  MoveL 3592 to (0, -43.6, 16.44) mm, rotated rx 90 ry 0 rz 180 deg; joints [1.406, -71.721, 106.574, -177.541, 34.877, 177.982]
  MoveL 3593 to (0, -43.6, 17.04) mm, rotated rx 90 ry 0 rz 180 deg; joints [1.381, -71.722, 106.575, -177.584, 34.877, 178.018]
  MoveL 3594 to (-200, -43.6, 17.04) mm, rotated rx 90 ry 0 rz 180 deg; joints [1.617, -84.213, 122.025, -177.364, 37.842, 177.918]
  MoveL 3595 to (-200, -43.6, 17.64) mm, rotated rx 90 ry 0 rz 180 deg; joints [1.587, -84.214, 122.026, -177.412, 37.841, 177.956]
  MoveL 3596 to (0, -43.6, 17.64) mm, rotated rx 90 ry 0 rz 180 deg; joints [1.356, -71.723, 106.576, -177.628, 34.876, 178.054]
  MoveL 3597 to (0, -43.6, 18.24) mm, rotated rx 90 ry 0 rz 180 deg; joints [1.331, -71.724, 106.577, -177.672, 34.876, 178.09]
  MoveL 3598 to (-200, -43.6, 18.24) mm, rotated rx 90 ry 0 rz 180 deg; joints [1.558, -84.215, 122.027, -177.46, 37.84, 177.993]
  MoveL 3599 to (-200, -43.6, 18.84) mm, rotated rx 90 ry 0 rz 180 deg; joints [1.529, -84.216, 122.028, -177.508, 37.839, 178.031]
  MoveL 3600 to (0, -43.6, 18.84) mm, rotated rx 90 ry 0 rz 180 deg; joints [1.306, -71.725, 106.578, -177.716, 34.875, 178.126]
  MoveL 3601 to (0, -43.6, 19.44) mm, rotated rx 90 ry 0 rz 180 deg; joints [1.281, -71.725, 106.579, -177.759, 34.875, 178.162]
  MoveL 3602 to (-200, -43.6, 19.44) mm, rotated rx 90 ry 0 rz 180 deg; joints [1.499, -84.217, 122.03, -177.555, 37.838, 178.069]
  MoveL 3603 to (-200, -43.6, 20.04) mm, rotated rx 90 ry 0 rz 180 deg; joints [1.47, -84.218, 122.031, -177.603, 37.837, 178.107]
  MoveL 3604 to (0, -43.6, 20.04) mm, rotated rx 90 ry 0 rz 180 deg; joints [1.256, -71.726, 106.58, -177.803, 34.874, 178.197]
  MoveL 3605 to (0, -43.6, 20.64) mm, rotated rx 90 ry 0 rz 180 deg; joints [1.231, -71.727, 106.582, -177.847, 34.874, 178.233]
  MoveL 3606 to (-200, -43.6, 20.64) mm, rotated rx 90 ry 0 rz 180 deg; joints [1.441, -84.219, 122.032, -177.651, 37.836, 178.144]
  MoveL 3607 to (-200, -43.6, 21.24) mm, rotated rx 90 ry 0 rz 180 deg; joints [1.411, -84.22, 122.033, -177.699, 37.835, 178.182]
  MoveL 3608 to (0, -43.6, 21.24) mm, rotated rx 90 ry 0 rz 180 deg; joints [1.206, -71.728, 106.583, -177.891, 34.873, 178.269]
  MoveL 3609 to (0, -43.6, 21.84) mm, rotated rx 90 ry 0 rz 180 deg; joints [1.181, -71.729, 106.584, -177.935, 34.873, 178.305]
  MoveL 3610 to (-200, -43.6, 21.84) mm, rotated rx 90 ry 0 rz 180 deg; joints [1.382, -84.221, 122.034, -177.746, 37.835, 178.22]
  MoveL 3611 to (-200, -43.6, 22.44) mm, rotated rx 90 ry 0 rz 180 deg; joints [1.353, -84.222, 122.035, -177.794, 37.834, 178.258]
  MoveL 3612 to (0, -43.6, 22.44) mm, rotated rx 90 ry 0 rz 180 deg; joints [1.156, -71.729, 106.585, -177.978, 34.872, 178.341]
  MoveL 3613 to (0, -43.6, 23.04) mm, rotated rx 90 ry 0 rz 180 deg; joints [1.131, -71.73, 106.586, -178.022, 34.872, 178.377]
  MoveL 3614 to (-200, -43.6, 23.04) mm, rotated rx 90 ry 0 rz 180 deg; joints [1.323, -84.223, 122.036, -177.842, 37.833, 178.295]
  MoveL 3615 to (-200, -43.6, 23.64) mm, rotated rx 90 ry 0 rz 180 deg; joints [1.294, -84.223, 122.037, -177.89, 37.832, 178.333]
  MoveL 3616 to (0, -43.6, 23.64) mm, rotated rx 90 ry 0 rz 180 deg; joints [1.106, -71.731, 106.587, -178.066, 34.871, 178.413]
  MoveL 3617 to (0, -43.6, 24.24) mm, rotated rx 90 ry 0 rz 180 deg; joints [1.081, -71.731, 106.588, -178.11, 34.871, 178.449]
  MoveL 3618 to (-200, -43.6, 24.24) mm, rotated rx 90 ry 0 rz 180 deg; joints [1.265, -84.224, 122.038, -177.938, 37.832, 178.371]
  MoveL 3619 to (-200, -43.6, 24.84) mm, rotated rx 90 ry 0 rz 180 deg; joints [1.236, -84.225, 122.039, -177.985, 37.831, 178.408]
  MoveL 3620 to (0, -43.6, 24.84) mm, rotated rx 90 ry 0 rz 180 deg; joints [1.055, -71.732, 106.589, -178.154, 34.87, 178.485]
  MoveL 3621 to (0, -43.6, 25.44) mm, rotated rx 90 ry 0 rz 180 deg; joints [1.03, -71.733, 106.589, -178.197, 34.87, 178.521]
  MoveL 3622 to (-200, -43.6, 25.44) mm, rotated rx 90 ry 0 rz 180 deg; joints [1.206, -84.226, 122.04, -178.033, 37.83, 178.446]
  MoveL 3623 to (-200, -43.6, 26.04) mm, rotated rx 90 ry 0 rz 180 deg; joints [1.177, -84.227, 122.041, -178.081, 37.829, 178.484]
  MoveL 3624 to (0, -43.6, 26.04) mm, rotated rx 90 ry 0 rz 180 deg; joints [1.005, -71.733, 106.59, -178.241, 34.87, 178.557]
  MoveL 3625 to (0, -43.6, 26.64) mm, rotated rx 90 ry 0 rz 180 deg; joints [0.98, -71.734, 106.591, -178.285, 34.869, 178.593]
  MoveL 3626 to (-200, -43.6, 26.64) mm, rotated rx 90 ry 0 rz 180 deg; joints [1.148, -84.228, 122.042, -178.129, 37.829, 178.522]
  MoveL 3627 to (-200, -43.6, 27.24) mm, rotated rx 90 ry 0 rz 180 deg; joints [1.118, -84.228, 122.042, -178.176, 37.828, 178.559]
  MoveL 3628 to (0, -43.6, 27.24) mm, rotated rx 90 ry 0 rz 180 deg; joints [0.955, -71.735, 106.592, -178.329, 34.869, 178.629]
  MoveL 3629 to (0, -43.6, 27.84) mm, rotated rx 90 ry 0 rz 180 deg; joints [0.93, -71.735, 106.593, -178.373, 34.868, 178.665]
  MoveL 3630 to (-200, -43.6, 27.84) mm, rotated rx 90 ry 0 rz 180 deg; joints [1.089, -84.229, 122.043, -178.224, 37.827, 178.597]
  MoveL 3631 to (-200, -43.6, 28.44) mm, rotated rx 90 ry 0 rz 180 deg; joints [1.06, -84.23, 122.044, -178.272, 37.827, 178.635]
  MoveL 3632 to (0, -43.6, 28.44) mm, rotated rx 90 ry 0 rz 180 deg; joints [0.905, -71.736, 106.594, -178.417, 34.868, 178.701]
  MoveL 3633 to (0, -43.6, 29.04) mm, rotated rx 90 ry 0 rz 180 deg; joints [0.88, -71.737, 106.594, -178.46, 34.868, 178.737]
  MoveL 3634 to (-200, -43.6, 29.04) mm, rotated rx 90 ry 0 rz 180 deg; joints [1.03, -84.23, 122.045, -178.32, 37.826, 178.673]
  MoveL 3635 to (-200, -43.6, 29.64) mm, rotated rx 90 ry 0 rz 180 deg; joints [1.001, -84.231, 122.046, -178.368, 37.826, 178.711]
  MoveL 3636 to (0, -43.6, 29.64) mm, rotated rx 90 ry 0 rz 180 deg; joints [0.855, -71.737, 106.595, -178.504, 34.867, 178.773]
  MoveL 3637 to (0, -43.6, 30.24) mm, rotated rx 90 ry 0 rz 180 deg; joints [0.83, -71.738, 106.596, -178.548, 34.867, 178.809]
  MoveL 3638 to (-200, -43.6, 30.24) mm, rotated rx 90 ry 0 rz 180 deg; joints [0.972, -84.232, 122.046, -178.416, 37.825, 178.748]
  MoveL 3639 to (-200, -43.6, 30.84) mm, rotated rx 90 ry 0 rz 180 deg; joints [0.942, -84.232, 122.047, -178.463, 37.825, 178.786]
  MoveL 3640 to (0, -43.6, 30.84) mm, rotated rx 90 ry 0 rz 180 deg; joints [0.805, -71.738, 106.597, -178.592, 34.867, 178.845]
  MoveL 3641 to (0, -43.6, 31.44) mm, rotated rx 90 ry 0 rz 180 deg; joints [0.78, -71.739, 106.597, -178.636, 34.866, 178.88]
  MoveL 3642 to (-200, -43.6, 31.44) mm, rotated rx 90 ry 0 rz 180 deg; joints [0.913, -84.233, 122.048, -178.511, 37.824, 178.824]
  MoveL 3643 to (-200, -43.6, 32.04) mm, rotated rx 90 ry 0 rz 180 deg; joints [0.884, -84.234, 122.048, -178.559, 37.823, 178.862]
  MoveL 3644 to (0, -43.6, 32.04) mm, rotated rx 90 ry 0 rz 180 deg; joints [0.755, -71.739, 106.598, -178.679, 34.866, 178.916]
  MoveL 3645 to (0, -43.6, 32.64) mm, rotated rx 90 ry 0 rz 180 deg; joints [0.73, -71.74, 106.599, -178.723, 34.866, 178.952]
  MoveL 3646 to (-200, -43.6, 32.64) mm, rotated rx 90 ry 0 rz 180 deg; joints [0.854, -84.234, 122.049, -178.607, 37.823, 178.899]
  MoveL 3647 to (-200, -43.6, 33.24) mm, rotated rx 90 ry 0 rz 180 deg; joints [0.825, -84.235, 122.05, -178.655, 37.822, 178.937]
  MoveL 3648 to (0, -43.6, 33.24) mm, rotated rx 90 ry 0 rz 180 deg; joints [0.705, -71.74, 106.599, -178.767, 34.865, 178.988]
  MoveL 3649 to (0, -43.6, 33.84) mm, rotated rx 90 ry 0 rz 180 deg; joints [0.68, -71.741, 106.6, -178.811, 34.865, 179.024]
  MoveL 3650 to (-200, -43.6, 33.84) mm, rotated rx 90 ry 0 rz 180 deg; joints [0.796, -84.235, 122.05, -178.702, 37.822, 178.975]
  MoveL 3651 to (-200, -43.6, 34.44) mm, rotated rx 90 ry 0 rz 180 deg; joints [0.766, -84.236, 122.051, -178.75, 37.822, 179.013]
  MoveL 3652 to (0, -43.6, 34.44) mm, rotated rx 90 ry 0 rz 180 deg; joints [0.655, -71.741, 106.6, -178.855, 34.865, 179.06]
  MoveL 3653 to (0, -43.6, 35.04) mm, rotated rx 90 ry 0 rz 180 deg; joints [0.63, -71.741, 106.601, -178.899, 34.865, 179.096]
  MoveL 3654 to (-200, -43.6, 35.04) mm, rotated rx 90 ry 0 rz 180 deg; joints [0.737, -84.236, 122.051, -178.798, 37.821, 179.05]
  MoveL 3655 to (-200, -43.6, 35.64) mm, rotated rx 90 ry 0 rz 180 deg; joints [0.708, -84.237, 122.052, -178.846, 37.821, 179.088]
  MoveL 3656 to (0, -43.6, 35.64) mm, rotated rx 90 ry 0 rz 180 deg; joints [0.605, -71.742, 106.602, -178.942, 34.864, 179.132]
  MoveL 3657 to (0, -43.6, 36.24) mm, rotated rx 90 ry 0 rz 180 deg; joints [0.579, -71.742, 106.602, -178.986, 34.864, 179.168]
  MoveL 3658 to (-200, -43.6, 36.24) mm, rotated rx 90 ry 0 rz 180 deg; joints [0.678, -84.237, 122.053, -178.894, 37.82, 179.126]
  MoveL 3659 to (-200, -43.6, 36.84) mm, rotated rx 90 ry 0 rz 180 deg; joints [0.649, -84.238, 122.053, -178.942, 37.82, 179.164]
  MoveL 3660 to (0, -43.6, 36.84) mm, rotated rx 90 ry 0 rz 180 deg; joints [0.554, -71.743, 106.603, -179.03, 34.864, 179.204]
  MoveL 3661 to (0, -43.6, 37.44) mm, rotated rx 90 ry 0 rz 180 deg; joints [0.529, -71.743, 106.603, -179.074, 34.864, 179.24]
  MoveL 3662 to (-200, -43.6, 37.44) mm, rotated rx 90 ry 0 rz 180 deg; joints [0.62, -84.238, 122.053, -178.989, 37.82, 179.202]
  MoveL 3663 to (-200, -43.6, 38.04) mm, rotated rx 90 ry 0 rz 180 deg; joints [0.59, -84.239, 122.054, -179.037, 37.819, 179.239]
  MoveL 3664 to (0, -43.6, 38.04) mm, rotated rx 90 ry 0 rz 180 deg; joints [0.504, -71.743, 106.603, -179.118, 34.863, 179.276]
  MoveL 3665 to (0, -43.6, 38.64) mm, rotated rx 90 ry 0 rz 180 deg; joints [0.479, -71.744, 106.604, -179.162, 34.863, 179.312]
  MoveL 3666 to (-200, -43.6, 38.64) mm, rotated rx 90 ry 0 rz 180 deg; joints [0.561, -84.239, 122.054, -179.085, 37.819, 179.277]
  MoveL 3667 to (-200, -43.6, 39.24) mm, rotated rx 90 ry 0 rz 180 deg; joints [0.532, -84.239, 122.055, -179.133, 37.819, 179.315]
  MoveL 3668 to (0, -43.6, 39.24) mm, rotated rx 90 ry 0 rz 180 deg; joints [0.454, -71.744, 106.604, -179.205, 34.863, 179.348]
  MoveL 3669 to (0, -43.6, 39.84) mm, rotated rx 90 ry 0 rz 180 deg; joints [0.429, -71.744, 106.605, -179.249, 34.863, 179.384]
  MoveL 3670 to (-200, -43.6, 39.84) mm, rotated rx 90 ry 0 rz 180 deg; joints [0.502, -84.24, 122.055, -179.181, 37.818, 179.353]
  MoveL 3671 to (-200, -43.6, 40.44) mm, rotated rx 90 ry 0 rz 180 deg; joints [0.473, -84.24, 122.056, -179.229, 37.818, 179.391]
  MoveL 3672 to (0, -43.6, 40.44) mm, rotated rx 90 ry 0 rz 180 deg; joints [0.404, -71.744, 106.605, -179.293, 34.863, 179.42]
  MoveL 3673 to (0, -43.6, 41.04) mm, rotated rx 90 ry 0 rz 180 deg; joints [0.379, -71.745, 106.605, -179.337, 34.863, 179.456]
  MoveL 3674 to (-200, -43.6, 41.04) mm, rotated rx 90 ry 0 rz 180 deg; joints [0.444, -84.24, 122.056, -179.276, 37.818, 179.428]
  MoveL 3675 to (-200, -43.6, 41.64) mm, rotated rx 90 ry 0 rz 180 deg; joints [0.414, -84.241, 122.056, -179.324, 37.817, 179.466]
  MoveL 3676 to (0, -43.6, 41.64) mm, rotated rx 90 ry 0 rz 180 deg; joints [0.354, -71.745, 106.606, -179.381, 34.862, 179.492]
  MoveL 3677 to (0, -43.6, 42.24) mm, rotated rx 90 ry 0 rz 180 deg; joints [0.329, -71.745, 106.606, -179.425, 34.862, 179.528]
  MoveL 3678 to (-200, -43.6, 42.24) mm, rotated rx 90 ry 0 rz 180 deg; joints [0.385, -84.241, 122.057, -179.372, 37.817, 179.504]
  MoveL 3679 to (-200, -43.6, 42.84) mm, rotated rx 90 ry 0 rz 180 deg; joints [0.356, -84.241, 122.057, -179.42, 37.817, 179.542]
  MoveL 3680 to (0, -43.6, 42.84) mm, rotated rx 90 ry 0 rz 180 deg; joints [0.304, -71.745, 106.606, -179.468, 34.862, 179.564]
  MoveL 3681 to (0, -43.6, 43.44) mm, rotated rx 90 ry 0 rz 180 deg; joints [0.279, -71.745, 106.607, -179.512, 34.862, 179.6]
  MoveL 3682 to (-200, -43.6, 43.44) mm, rotated rx 90 ry 0 rz 180 deg; joints [0.326, -84.241, 122.057, -179.468, 37.817, 179.579]
  MoveL 3683 to (-200, -43.6, 44.04) mm, rotated rx 90 ry 0 rz 180 deg; joints [0.297, -84.242, 122.057, -179.516, 37.817, 179.617]
  MoveL 3684 to (0, -43.6, 44.04) mm, rotated rx 90 ry 0 rz 180 deg; joints [0.254, -71.746, 106.607, -179.556, 34.862, 179.636]
  MoveL 3685 to (0, -43.6, 44.64) mm, rotated rx 90 ry 0 rz 180 deg; joints [0.229, -71.746, 106.607, -179.6, 34.862, 179.672]
  MoveL 3686 to (-200, -43.6, 44.64) mm, rotated rx 90 ry 0 rz 180 deg; joints [0.268, -84.242, 122.057, -179.563, 37.816, 179.655]
  MoveL 3687 to (-200, -43.6, 45.24) mm, rotated rx 91 ry 0 rz 180 deg; joints [-0.066, -84.215, 122.091, 179.892, 37.876, -178.916]
  MoveL 3688 to (0, -43.6, 45.24) mm, rotated rx 91 ry 0 rz 180 deg; joints [-0.057, -71.723, 106.638, 179.901, 34.915, -178.92]
  MoveL 3689 to (0, -43.57, 45.84) mm, rotated rx 93.53 ry 0 rz 180 deg; joints [-0.737, -71.643, 106.723, 178.718, 35.087, -175.424]
  MoveL 3690 to (-200, -43.57, 45.84) mm, rotated rx 93.53 ry 0 rz 180 deg; joints [-0.863, -84.12, 122.183, 178.601, 38.071, -175.372]
  MoveL 3691 to (-200, -43.52, 46.43) mm, rotated rx 96.06 ry 0 rz 180 deg; joints [-1.652, -83.985, 122.287, 177.335, 38.332, -171.854]
  MoveL 3692 to (0, -43.52, 46.43) mm, rotated rx 96.06 ry 0 rz 180 deg; joints [-1.412, -71.53, 106.819, 177.558, 35.313, -171.952]
  MoveL 3693 to (0, -43.45, 47.03) mm, rotated rx 98.58 ry 0 rz 180 deg; joints [-2.079, -71.385, 106.923, 176.426, 35.591, -168.511]
  MoveL 3694 to (-200, -43.45, 47.03) mm, rotated rx 98.58 ry 0 rz 180 deg; joints [-2.433, -83.81, 122.402, 176.102, 38.656, -168.373]
  MoveL 3695 to (-200, -43.34, 47.62) mm, rotated rx 101.11 ry 0 rz 180 deg; joints [-3.205, -83.596, 122.528, 174.908, 39.042, -164.931]
  MoveL 3696 to (0, -43.34, 47.62) mm, rotated rx 101.11 ry 0 rz 180 deg; joints [-2.738, -71.207, 107.038, 175.329, 35.922, -165.105]
  MoveL 3697 to (0, -43.22, 48.21) mm, rotated rx 103.64 ry 0 rz 180 deg; joints [-3.387, -70.996, 107.161, 174.272, 36.301, -161.74]
  MoveL 3698 to (-200, -43.22, 48.21) mm, rotated rx 103.64 ry 0 rz 180 deg; joints [-3.964, -83.344, 122.664, 173.759, 39.488, -161.538]
  MoveL 3699 to (-200, -43.06, 48.79) mm, rotated rx 106.17 ry 0 rz 180 deg; joints [-4.709, -83.052, 122.811, 172.66, 39.991, -158.198]
  MoveL 3700 to (0, -43.06, 48.79) mm, rotated rx 106.17 ry 0 rz 180 deg; joints [-4.025, -70.753, 107.292, 173.259, 36.729, -158.423]
  MoveL 3701 to (0, -42.88, 49.36) mm, rotated rx 108.69 ry 0 rz 180 deg; joints [-4.65, -70.479, 107.431, 172.294, 37.203, -155.156]
  MoveL 3702 to (-200, -42.88, 49.36) mm, rotated rx 108.69 ry 0 rz 180 deg; joints [-5.439, -82.722, 122.966, 171.616, 40.548, -154.917]
  MoveL 3703 to (-200, -42.68, 49.92) mm, rotated rx 111.22 ry 0 rz 180 deg; joints [-6.153, -82.354, 123.131, 170.627, 41.159, -151.695]
  MoveL 3704 to (0, -42.68, 49.92) mm, rotated rx 111.22 ry 0 rz 180 deg; joints [-5.261, -70.173, 107.578, 171.38, 37.72, -151.941]
  MoveL 3705 to (0, -42.45, 50.48) mm, rotated rx 113.75 ry 0 rz 180 deg; joints [-5.857, -69.835, 107.731, 170.518, 38.278, -148.781]
  MoveL 3706 to (-200, -42.45, 50.48) mm, rotated rx 113.75 ry 0 rz 180 deg; joints [-6.848, -81.948, 123.304, 169.698, 41.818, -148.537]
  MoveL 3707 to (-200, -42.2, 51.02) mm, rotated rx 116.28 ry 0 rz 180 deg; joints [-7.524, -81.505, 123.483, 168.83, 42.524, -145.443]
  MoveL 3708 to (0, -42.2, 51.02) mm, rotated rx 116.28 ry 0 rz 180 deg; joints [-6.437, -69.468, 107.89, 169.711, 38.876, -145.679]
  MoveL 3709 to (0, -41.92, 51.55) mm, rotated rx 118.8 ry 0 rz 180 deg; joints [-6.999, -69.07, 108.055, 168.959, 39.51, -142.635]
  MoveL 3710 to (-200, -41.92, 51.55) mm, rotated rx 118.8 ry 0 rz 180 deg; joints [-8.178, -81.025, 123.67, 168.023, 43.273, -142.416]
  MoveL 3711 to (-200, -41.62, 52.07) mm, rotated rx 121.33 ry 0 rz 180 deg; joints [-8.81, -80.51, 123.862, 167.278, 44.064, -139.453]
  MoveL 3712 to (0, -41.62, 52.07) mm, rotated rx 121.33 ry 0 rz 180 deg; joints [-7.542, -68.643, 108.225, 168.262, 40.178, -139.647]
  MoveL 3713 to (0, -41.29, 52.58) mm, rotated rx 123.86 ry 0 rz 180 deg; joints [-8.065, -68.186, 108.399, 167.621, 40.878, -136.717]
  MoveL 3714 to (-200, -41.29, 52.58) mm, rotated rx 123.86 ry 0 rz 180 deg; joints [-9.419, -79.959, 124.059, 166.593, 44.892, -136.555]
  MoveL 3715 to (-200, -40.95, 53.07) mm, rotated rx 126.39 ry 0 rz 180 deg; joints [-10.003, -79.373, 124.26, 165.967, 45.755, -133.72]
  MoveL 3716 to (0, -40.95, 53.07) mm, rotated rx 126.39 ry 0 rz 180 deg; joints [-8.568, -67.702, 108.576, 167.034, 41.607, -133.844]
  MoveL 3717 to (0, -40.58, 53.54) mm, rotated rx 128.92 ry 0 rz 180 deg; joints [-9.05, -67.19, 108.755, 166.501, 42.364, -131.026]
  MoveL 3718 to (-200, -40.58, 53.54) mm, rotated rx 128.92 ry 0 rz 180 deg; joints [-10.562, -78.754, 124.464, 165.4, 46.65, -130.946]
  MoveL 3719 to (-200, -40.2, 54) mm, rotated rx 131.44 ry 0 rz 180 deg; joints [-11.094, -78.102, 124.671, 164.89, 47.574, -128.233]
  MoveL 3720 to (0, -40.2, 54) mm, rotated rx 131.44 ry 0 rz 180 deg; joints [-9.508, -66.651, 108.937, 166.021, 43.144, -128.262]
  MoveL 3721 to (0, -39.79, 54.44) mm, rotated rx 133.97 ry 0 rz 180 deg; joints [-9.944, -66.086, 109.12, 165.592, 43.948, -125.549]
  MoveL 3722 to (-200, -39.79, 54.44) mm, rotated rx 133.97 ry 0 rz 180 deg; joints [-11.599, -77.418, 124.879, 164.435, 48.526, -125.576]
  MoveL 3723 to (-200, -39.36, 54.87) mm, rotated rx 136.5 ry 0 rz 180 deg; joints [-12.075, -76.703, 125.088, 164.032, 49.502, -122.974]
  MoveL 3724 to (0, -39.36, 54.87) mm, rotated rx 136.5 ry 0 rz 180 deg; joints [-10.356, -65.497, 109.304, 165.212, 44.772, -122.886]
  MoveL 3725 to (0, -38.92, 55.27) mm, rotated rx 139.03 ry 0 rz 180 deg; joints [-10.744, -64.883, 109.487, 164.879, 45.614, -120.27]
  MoveL 3726 to (-200, -38.92, 55.27) mm, rotated rx 139.03 ry 0 rz 180 deg; joints [-12.523, -75.959, 125.297, 163.679, 50.5, -120.422]
  MoveL 3727 to (-200, -38.46, 55.65) mm, rotated rx 141.55 ry 0 rz 180 deg; joints [-12.942, -75.185, 125.505, 163.375, 51.517, -117.92]
  MoveL 3728 to (0, -38.46, 55.65) mm, rotated rx 141.55 ry 0 rz 180 deg; joints [-11.106, -64.246, 109.67, 164.593, 46.471, -117.699]
  MoveL 3729 to (0, -37.98, 56.01) mm, rotated rx 144.08 ry 0 rz 180 deg; joints [-11.442, -63.587, 109.851, 164.351, 47.344, -115.17]
  MoveL 3730 to (-200, -37.98, 56.01) mm, rotated rx 144.08 ry 0 rz 180 deg; joints [-13.33, -74.384, 125.711, 163.117, 52.552, -115.462]
  MoveL 3731 to (-200, -37.48, 56.35) mm, rotated rx 146.61 ry 0 rz 180 deg; joints [-13.688, -73.557, 125.915, 162.903, 53.603, -113.047]
  MoveL 3732 to (0, -37.48, 56.35) mm, rotated rx 146.61 ry 0 rz 180 deg; joints [-11.753, -62.906, 110.029, 164.15, 48.228, -112.68]
  MoveL 3733 to (0, -36.98, 56.67) mm, rotated rx 149.14 ry 0 rz 180 deg; joints [-12.037, -62.206, 110.205, 163.99, 49.123, -110.227]
  MoveL 3734 to (-200, -36.98, 56.67) mm, rotated rx 149.14 ry 0 rz 180 deg; joints [-14.015, -72.704, 126.115, 162.731, 54.667, -110.67]
  MoveL 3735 to (-200, -36.45, 56.97) mm, rotated rx 151.66 ry 0 rz 180 deg; joints [-14.311, -71.828, 126.31, 162.598, 55.742, -108.329]
  MoveL 3736 to (0, -36.45, 56.97) mm, rotated rx 151.66 ry 0 rz 180 deg; joints [-12.293, -61.487, 110.377, 163.869, 50.027, -107.809]
  MoveL 3737 to (0, -35.92, 57.24) mm, rotated rx 154.19 ry 0 rz 180 deg; joints [-12.522, -60.751, 110.546, 163.785, 50.937, -105.422]
  MoveL 3738 to (-200, -35.92, 57.24) mm, rotated rx 154.19 ry 0 rz 180 deg; joints [-14.575, -70.93, 126.501, 162.504, 56.826, -106.021]
  MoveL 3739 to (-200, -35.38, 57.49) mm, rotated rx 156.72 ry 0 rz 180 deg; joints [-14.807, -70.01, 126.687, 162.445, 57.919, -103.741]
  MoveL 3740 to (0, -35.38, 57.49) mm, rotated rx 156.72 ry 0 rz 180 deg; joints [-12.724, -59.998, 110.709, 163.736, 51.853, -103.064]
  MoveL 3741 to (0, -34.82, 57.72) mm, rotated rx 159.25 ry 0 rz 180 deg; joints [-12.898, -59.23, 110.867, 163.72, 52.773, -100.732]
  MoveL 3742 to (-200, -34.82, 57.72) mm, rotated rx 159.25 ry 0 rz 180 deg; joints [-15.006, -69.072, 126.866, 162.421, 59.017, -101.488]
  MoveL 3743 to (-200, -34.25, 57.92) mm, rotated rx 161.78 ry 0 rz 180 deg; joints [-15.173, -68.116, 127.038, 162.43, 60.118, -99.259]
  MoveL 3744 to (0, -34.25, 57.92) mm, rotated rx 161.78 ry 0 rz 180 deg; joints [-13.043, -58.449, 111.02, 163.737, 53.694, -98.424]
  MoveL 3745 to (0, -33.68, 58.09) mm, rotated rx 164.3 ry 0 rz 180 deg; joints [-13.16, -57.655, 111.167, 163.784, 54.617, -96.137]
  MoveL 3746 to (-200, -33.68, 58.09) mm, rotated rx 164.3 ry 0 rz 180 deg; joints [-15.308, -67.145, 127.203, 162.47, 61.223, -97.05]
  MoveL 3747 to (-200, -33.1, 58.24) mm, rotated rx 166.83 ry 0 rz 180 deg; joints [-15.409, -66.159, 127.36, 162.54, 62.327, -94.858]
  MoveL 3748 to (0, -33.1, 58.24) mm, rotated rx 166.83 ry 0 rz 180 deg; joints [-13.249, -56.85, 111.306, 163.862, 55.538, -93.869]
  MoveL 3749 to (0, -32.51, 58.37) mm, rotated rx 169.36 ry 0 rz 180 deg; joints [-13.308, -56.037, 111.439, 163.967, 56.458, -91.618]
  MoveL 3750 to (-200, -32.51, 58.37) mm, rotated rx 169.36 ry 0 rz 180 deg; joints [-15.478, -65.161, 127.509, 162.64, 63.431, -92.68]
  MoveL 3751 to (-200, -31.92, 58.46) mm, rotated rx 171.89 ry 0 rz 180 deg; joints [-15.514, -64.153, 127.649, 162.767, 64.532, -90.516]
  MoveL 3752 to (0, -31.92, 58.46) mm, rotated rx 171.89 ry 0 rz 180 deg; joints [-13.34, -55.215, 111.565, 164.1, 57.373, -89.382]
  MoveL 3753 to (0, -31.32, 58.53) mm, rotated rx 174.41 ry 0 rz 180 deg; joints [-13.342, -54.388, 111.683, 164.26, 58.283, -87.157]
  MoveL 3754 to (-200, -31.32, 58.53) mm, rotated rx 174.41 ry 0 rz 180 deg; joints [-15.517, -63.136, 127.779, 162.921, 65.629, -88.36]
  MoveL 3755 to (-200, -30.73, 58.58) mm, rotated rx 176.94 ry 0 rz 180 deg; joints [-15.486, -62.113, 127.901, 163.102, 66.72, -86.21]
  MoveL 3756 to (0, -30.73, 58.58) mm, rotated rx 176.94 ry 0 rz 180 deg; joints [-13.316, -53.555, 111.794, 164.445, 59.187, -84.942]
  MoveL 3757 to (0, -30.13, 58.6) mm, rotated rx 179.47 ry 0 rz 180 deg; joints [-13.261, -52.72, 111.896, 164.654, 60.083, -82.735]
  MoveL 3758 to (-200, -30.13, 58.6) mm, rotated rx 179.47 ry 0 rz 180 deg; joints [-15.423, -61.085, 128.012, 163.308, 67.803, -84.066]
  MoveL 3759 to (-200, -29.53, 58.6) mm, rotated rx 180 ry 0 rz 180 deg; joints [-15.406, -60.839, 128.036, 163.358, 68.06, -83.627]
  MoveL 3760 to (0, -29.53, 58.6) mm, rotated rx 180 ry 0 rz 180 deg; joints [-13.245, -52.52, 111.918, 164.705, 60.295, -82.283]
  MoveL 3761 to (0, -28.93, 58.6) mm, rotated rx 180 ry 0 rz 180 deg; joints [-13.245, -52.489, 111.92, 164.71, 60.328, -82.293]
  MoveL 3762 to (-200, -28.93, 58.6) mm, rotated rx 180 ry 0 rz 180 deg; joints [-15.406, -60.801, 128.039, 163.362, 68.099, -83.64]
  MoveL 3763 to (-200, -28.33, 58.6) mm, rotated rx 180 ry 0 rz 180 deg; joints [-15.406, -60.762, 128.041, 163.367, 68.138, -83.652]
  MoveL 3764 to (0, -28.33, 58.6) mm, rotated rx 180 ry 0 rz 180 deg; joints [-13.245, -52.457, 111.922, 164.715, 60.36, -82.303]
  MoveL 3765 to (0, -27.73, 58.6) mm, rotated rx 180 ry 0 rz 180 deg; joints [-13.245, -52.426, 111.924, 164.72, 60.392, -82.313]
  MoveL 3766 to (-200, -27.73, 58.6) mm, rotated rx 180 ry 0 rz 180 deg; joints [-15.406, -60.724, 128.043, 163.372, 68.177, -83.665]
  MoveL 3767 to (-200, -27.13, 58.6) mm, rotated rx 180 ry 0 rz 180 deg; joints [-15.406, -60.685, 128.046, 163.377, 68.216, -83.678]
  MoveL 3768 to (0, -27.13, 58.6) mm, rotated rx 180 ry 0 rz 180 deg; joints [-13.245, -52.395, 111.926, 164.725, 60.424, -82.323]
  MoveL 3769 to (0, -26.53, 58.6) mm, rotated rx 180 ry 0 rz 180 deg; joints [-13.245, -52.363, 111.928, 164.73, 60.457, -82.333]
  MoveL 3770 to (-200, -26.53, 58.6) mm, rotated rx 180 ry 0 rz 180 deg; joints [-15.406, -60.647, 128.048, 163.381, 68.255, -83.69]
  MoveL 3771 to (-200, -25.93, 58.6) mm, rotated rx 180 ry 0 rz 180 deg; joints [-15.406, -60.608, 128.05, 163.386, 68.294, -83.703]
  MoveL 3772 to (0, -25.93, 58.6) mm, rotated rx 180 ry 0 rz 180 deg; joints [-13.245, -52.332, 111.93, 164.735, 60.489, -82.343]
  MoveL 3773 to (0, -25.33, 58.6) mm, rotated rx 180 ry 0 rz 180 deg; joints [-13.245, -52.3, 111.932, 164.74, 60.521, -82.354]
  MoveL 3774 to (-200, -25.33, 58.6) mm, rotated rx 180 ry 0 rz 180 deg; joints [-15.406, -60.57, 128.052, 163.39, 68.333, -83.715]
  MoveL 3775 to (-200, -24.73, 58.6) mm, rotated rx 180 ry 0 rz 180 deg; joints [-15.406, -60.531, 128.054, 163.395, 68.372, -83.728]
  MoveL 3776 to (0, -24.73, 58.6) mm, rotated rx 180 ry 0 rz 180 deg; joints [-13.245, -52.269, 111.934, 164.745, 60.553, -82.364]
  MoveL 3777 to (0, -24.13, 58.6) mm, rotated rx 180 ry 0 rz 180 deg; joints [-13.245, -52.237, 111.936, 164.75, 60.585, -82.374]
  MoveL 3778 to (-200, -24.13, 58.6) mm, rotated rx 180 ry 0 rz 180 deg; joints [-15.406, -60.492, 128.056, 163.4, 68.411, -83.74]
  MoveL 3779 to (-200, -23.53, 58.6) mm, rotated rx 180 ry 0 rz 180 deg; joints [-15.406, -60.454, 128.058, 163.404, 68.45, -83.753]
  MoveL 3780 to (0, -23.53, 58.6) mm, rotated rx 180 ry 0 rz 180 deg; joints [-13.245, -52.206, 111.938, 164.755, 60.618, -82.384]
  MoveL 3781 to (0, -22.93, 58.6) mm, rotated rx 180 ry 0 rz 180 deg; joints [-13.245, -52.174, 111.939, 164.76, 60.65, -82.394]
  MoveL 3782 to (-200, -22.93, 58.6) mm, rotated rx 180 ry 0 rz 180 deg; joints [-15.406, -60.415, 128.06, 163.409, 68.489, -83.765]
  MoveL 3783 to (-200, -22.33, 58.6) mm, rotated rx 180 ry 0 rz 180 deg; joints [-15.406, -60.376, 128.062, 163.413, 68.528, -83.778]
  MoveL 3784 to (0, -22.33, 58.6) mm, rotated rx 180 ry 0 rz 180 deg; joints [-13.245, -52.143, 111.941, 164.765, 60.682, -82.404]
  MoveL 3785 to (0, -21.73, 58.6) mm, rotated rx 180 ry 0 rz 180 deg; joints [-13.245, -52.111, 111.943, 164.77, 60.714, -82.414]
  MoveL 3786 to (-200, -21.73, 58.6) mm, rotated rx 180 ry 0 rz 180 deg; joints [-15.406, -60.338, 128.064, 163.418, 68.567, -83.79]
  MoveL 3787 to (-200, -21.13, 58.6) mm, rotated rx 180 ry 0 rz 180 deg; joints [-15.406, -60.299, 128.066, 163.423, 68.606, -83.803]
  MoveL 3788 to (0, -21.13, 58.6) mm, rotated rx 180 ry 0 rz 180 deg; joints [-13.245, -52.079, 111.945, 164.775, 60.746, -82.424]
  MoveL 3789 to (0, -20.53, 58.6) mm, rotated rx 180 ry 0 rz 180 deg; joints [-13.245, -52.048, 111.946, 164.78, 60.778, -82.434]
  MoveL 3790 to (-200, -20.53, 58.6) mm, rotated rx 180 ry 0 rz 180 deg; joints [-15.406, -60.26, 128.068, 163.427, 68.645, -83.815]
  MoveL 3791 to (-200, -19.93, 58.6) mm, rotated rx 180 ry 0 rz 180 deg; joints [-15.406, -60.221, 128.07, 163.432, 68.684, -83.828]
  MoveL 3792 to (0, -19.93, 58.6) mm, rotated rx 180 ry 0 rz 180 deg; joints [-13.245, -52.016, 111.948, 164.784, 60.81, -82.444]
  MoveL 3793 to (0, -19.33, 58.6) mm, rotated rx 180 ry 0 rz 180 deg; joints [-13.245, -51.985, 111.95, 164.789, 60.842, -82.454]
  MoveL 3794 to (-200, -19.33, 58.6) mm, rotated rx 180 ry 0 rz 180 deg; joints [-15.406, -60.182, 128.071, 163.436, 68.723, -83.84]
  MoveL 3795 to (-200, -18.73, 58.6) mm, rotated rx 180 ry 0 rz 180 deg; joints [-15.406, -60.144, 128.073, 163.441, 68.762, -83.852]
  MoveL 3796 to (0, -18.73, 58.6) mm, rotated rx 180 ry 0 rz 180 deg; joints [-13.245, -51.953, 111.951, 164.794, 60.874, -82.464]
  MoveL 3797 to (0, -18.13, 58.6) mm, rotated rx 180 ry 0 rz 180 deg; joints [-13.245, -51.921, 111.953, 164.799, 60.907, -82.474]
  MoveL 3798 to (-200, -18.13, 58.6) mm, rotated rx 180 ry 0 rz 180 deg; joints [-15.406, -60.105, 128.075, 163.445, 68.801, -83.865]
  MoveL 3799 to (-200, -17.53, 58.6) mm, rotated rx 180 ry 0 rz 180 deg; joints [-15.406, -60.066, 128.077, 163.45, 68.84, -83.877]
  MoveL 3800 to (0, -17.53, 58.6) mm, rotated rx 180 ry 0 rz 180 deg; joints [-13.245, -51.89, 111.954, 164.804, 60.939, -82.484]
  MoveL 3801 to (0, -16.93, 58.6) mm, rotated rx 180 ry 0 rz 180 deg; joints [-13.245, -51.858, 111.956, 164.809, 60.971, -82.494]
  MoveL 3802 to (-200, -16.93, 58.6) mm, rotated rx 180 ry 0 rz 180 deg; joints [-15.406, -60.027, 128.078, 163.454, 68.878, -83.89]
  MoveL 3803 to (-200, -16.33, 58.6) mm, rotated rx 180 ry 0 rz 180 deg; joints [-15.406, -59.988, 128.08, 163.458, 68.917, -83.902]
  MoveL 3804 to (0, -16.33, 58.6) mm, rotated rx 180 ry 0 rz 180 deg; joints [-13.245, -51.826, 111.957, 164.814, 61.003, -82.504]
  MoveL 3805 to (0, -15.73, 58.6) mm, rotated rx 180 ry 0 rz 180 deg; joints [-13.245, -51.795, 111.959, 164.818, 61.035, -82.514]
  MoveL 3806 to (-200, -15.73, 58.6) mm, rotated rx 180 ry 0 rz 180 deg; joints [-15.406, -59.949, 128.082, 163.463, 68.956, -83.914]
  MoveL 3807 to (-200, -15.13, 58.6) mm, rotated rx 180 ry 0 rz 180 deg; joints [-15.406, -59.91, 128.083, 163.467, 68.995, -83.927]
  MoveL 3808 to (0, -15.13, 58.6) mm, rotated rx 180 ry 0 rz 180 deg; joints [-13.245, -51.763, 111.96, 164.823, 61.067, -82.524]
  MoveL 3809 to (0, -14.53, 58.6) mm, rotated rx 180 ry 0 rz 180 deg; joints [-13.245, -51.731, 111.962, 164.828, 61.099, -82.534]
  MoveL 3810 to (-200, -14.53, 58.6) mm, rotated rx 180 ry 0 rz 180 deg; joints [-15.406, -59.871, 128.085, 163.472, 69.034, -83.939]
  MoveL 3811 to (-200, -13.93, 58.6) mm, rotated rx 180 ry 0 rz 180 deg; joints [-15.406, -59.833, 128.086, 163.476, 69.073, -83.951]
  MoveL 3812 to (0, -13.93, 58.6) mm, rotated rx 180 ry 0 rz 180 deg; joints [-13.245, -51.699, 111.963, 164.833, 61.131, -82.543]
  MoveL 3813 to (0, -13.33, 58.6) mm, rotated rx 180 ry 0 rz 180 deg; joints [-13.245, -51.667, 111.964, 164.838, 61.163, -82.553]
  MoveL 3814 to (-200, -13.33, 58.6) mm, rotated rx 180 ry 0 rz 180 deg; joints [-15.406, -59.794, 128.088, 163.481, 69.111, -83.964]
  MoveL 3815 to (-200, -12.73, 58.6) mm, rotated rx 180 ry 0 rz 180 deg; joints [-15.406, -59.755, 128.089, 163.485, 69.15, -83.976]
  MoveL 3816 to (0, -12.73, 58.6) mm, rotated rx 180 ry 0 rz 180 deg; joints [-13.245, -51.636, 111.966, 164.842, 61.194, -82.563]
  MoveL 3817 to (0, -12.13, 58.6) mm, rotated rx 180 ry 0 rz 180 deg; joints [-13.245, -51.604, 111.967, 164.847, 61.226, -82.573]
  MoveL 3818 to (-200, -12.13, 58.6) mm, rotated rx 180 ry 0 rz 180 deg; joints [-15.406, -59.716, 128.09, 163.489, 69.189, -83.988]
  MoveL 3819 to (-200, -11.53, 58.6) mm, rotated rx 180 ry 0 rz 180 deg; joints [-15.406, -59.677, 128.092, 163.494, 69.228, -84]
  MoveL 3820 to (0, -11.53, 58.6) mm, rotated rx 180 ry 0 rz 180 deg; joints [-13.245, -51.572, 111.968, 164.852, 61.258, -82.583]
  MoveL 3821 to (0, -10.93, 58.6) mm, rotated rx 180 ry 0 rz 180 deg; joints [-13.245, -51.54, 111.969, 164.857, 61.29, -82.593]
  MoveL 3822 to (-200, -10.93, 58.6) mm, rotated rx 180 ry 0 rz 180 deg; joints [-15.406, -59.637, 128.093, 163.498, 69.266, -84.013]
  MoveL 3823 to (-200, -10.33, 58.6) mm, rotated rx 180 ry 0 rz 180 deg; joints [-15.406, -59.598, 128.094, 163.502, 69.305, -84.025]
  MoveL 3824 to (0, -10.33, 58.6) mm, rotated rx 180 ry 0 rz 180 deg; joints [-13.245, -51.508, 111.97, 164.861, 61.322, -82.603]
  MoveL 3825 to (0, -9.73, 58.6) mm, rotated rx 180 ry 0 rz 180 deg; joints [-13.245, -51.476, 111.972, 164.866, 61.354, -82.612]
  MoveL 3826 to (-200, -9.73, 58.6) mm, rotated rx 180 ry 0 rz 180 deg; joints [-15.406, -59.559, 128.096, 163.507, 69.344, -84.037]
  MoveL 3827 to (-200, -9.13, 58.6) mm, rotated rx 180 ry 0 rz 180 deg; joints [-15.406, -59.52, 128.097, 163.511, 69.382, -84.049]
  MoveL 3828 to (0, -9.13, 58.6) mm, rotated rx 180 ry 0 rz 180 deg; joints [-13.245, -51.445, 111.973, 164.871, 61.386, -82.622]
  MoveL 3829 to (0, -8.53, 58.6) mm, rotated rx 180 ry 0 rz 180 deg; joints [-13.245, -51.413, 111.974, 164.875, 61.418, -82.632]
  MoveL 3830 to (-200, -8.53, 58.6) mm, rotated rx 180 ry 0 rz 180 deg; joints [-15.406, -59.481, 128.098, 163.515, 69.421, -84.062]
  MoveL 3831 to (-200, -7.93, 58.6) mm, rotated rx 180 ry 0 rz 180 deg; joints [-15.406, -59.442, 128.099, 163.52, 69.46, -84.074]
  MoveL 3832 to (0, -7.93, 58.6) mm, rotated rx 180 ry 0 rz 180 deg; joints [-13.245, -51.381, 111.975, 164.88, 61.45, -82.642]
  MoveL 3833 to (0, -7.33, 58.6) mm, rotated rx 180 ry 0 rz 180 deg; joints [-13.245, -51.349, 111.976, 164.885, 61.481, -82.652]
  MoveL 3834 to (-200, -7.33, 58.6) mm, rotated rx 180 ry 0 rz 180 deg; joints [-15.406, -59.403, 128.101, 163.524, 69.498, -84.086]
  MoveL 3835 to (-200, -6.73, 58.6) mm, rotated rx 180 ry 0 rz 180 deg; joints [-15.406, -59.364, 128.102, 163.528, 69.537, -84.098]
  MoveL 3836 to (0, -6.73, 58.6) mm, rotated rx 180 ry 0 rz 180 deg; joints [-13.245, -51.317, 111.977, 164.889, 61.513, -82.661]
  MoveL 3837 to (0, -6.13, 58.6) mm, rotated rx 180 ry 0 rz 180 deg; joints [-13.245, -51.285, 111.978, 164.894, 61.545, -82.671]
  MoveL 3838 to (-200, -6.13, 58.6) mm, rotated rx 180 ry 0 rz 180 deg; joints [-15.406, -59.325, 128.103, 163.532, 69.575, -84.11]
  MoveL 3839 to (-200, -5.53, 58.6) mm, rotated rx 180 ry 0 rz 180 deg; joints [-15.406, -59.285, 128.104, 163.537, 69.614, -84.123]
  MoveL 3840 to (0, -5.53, 58.6) mm, rotated rx 180 ry 0 rz 180 deg; joints [-13.245, -51.253, 111.979, 164.899, 61.577, -82.681]
  MoveL 3841 to (0, -4.93, 58.6) mm, rotated rx 180 ry 0 rz 180 deg; joints [-13.245, -51.221, 111.98, 164.903, 61.608, -82.691]
  MoveL 3842 to (-200, -4.93, 58.6) mm, rotated rx 180 ry 0 rz 180 deg; joints [-15.406, -59.246, 128.105, 163.541, 69.653, -84.135]
  MoveL 3843 to (-200, -4.33, 58.6) mm, rotated rx 180 ry 0 rz 180 deg; joints [-15.406, -59.207, 128.106, 163.545, 69.691, -84.147]
  MoveL 3844 to (0, -4.33, 58.6) mm, rotated rx 180 ry 0 rz 180 deg; joints [-13.245, -51.189, 111.981, 164.908, 61.64, -82.7]
  MoveL 3845 to (0, -3.73, 58.6) mm, rotated rx 180 ry 0 rz 180 deg; joints [-13.245, -51.157, 111.981, 164.913, 61.672, -82.71]
  MoveL 3846 to (-200, -3.73, 58.6) mm, rotated rx 180 ry 0 rz 180 deg; joints [-15.406, -59.168, 128.107, 163.549, 69.73, -84.159]
  MoveL 3847 to (-200, -3.13, 58.6) mm, rotated rx 180 ry 0 rz 180 deg; joints [-15.406, -59.128, 128.108, 163.553, 69.768, -84.171]
  MoveL 3848 to (0, -3.13, 58.6) mm, rotated rx 180 ry 0 rz 180 deg; joints [-13.245, -51.125, 111.982, 164.917, 61.704, -82.72]
  MoveL 3849 to (0, -2.53, 58.6) mm, rotated rx 180 ry 0 rz 180 deg; joints [-13.245, -51.093, 111.983, 164.922, 61.735, -82.73]
  MoveL 3850 to (-200, -2.53, 58.6) mm, rotated rx 180 ry 0 rz 180 deg; joints [-15.406, -59.089, 128.108, 163.558, 69.807, -84.183]
  MoveL 3851 to (-200, -1.93, 58.6) mm, rotated rx 180 ry 0 rz 180 deg; joints [-15.406, -59.05, 128.109, 163.562, 69.845, -84.195]
  MoveL 3852 to (0, -1.93, 58.6) mm, rotated rx 180 ry 0 rz 180 deg; joints [-13.245, -51.061, 111.984, 164.926, 61.767, -82.739]
  MoveL 3853 to (0, -1.33, 58.6) mm, rotated rx 180 ry 0 rz 180 deg; joints [-13.245, -51.029, 111.984, 164.931, 61.799, -82.749]
  MoveL 3854 to (-200, -1.33, 58.6) mm, rotated rx 180 ry 0 rz 180 deg; joints [-15.406, -59.01, 128.11, 163.566, 69.884, -84.207]
  MoveL 3855 to (-200, -0.73, 58.6) mm, rotated rx 180 ry 0 rz 180 deg; joints [-15.406, -58.971, 128.111, 163.57, 69.922, -84.22]
  MoveL 3856 to (0, -0.73, 58.6) mm, rotated rx 180 ry 0 rz 180 deg; joints [-13.245, -50.997, 111.985, 164.935, 61.83, -82.759]
  MoveL 3857 to (0, -0.13, 58.6) mm, rotated rx 180 ry 0 rz 180 deg; joints [-13.245, -50.964, 111.986, 164.94, 61.862, -82.768]
  MoveL 3858 to (-200, -0.13, 58.6) mm, rotated rx 180 ry 0 rz 180 deg; joints [-15.406, -58.932, 128.112, 163.574, 69.961, -84.232]
  MoveL 3859 to (-200, 0, 58.6) mm, rotated rx 180 ry 0 rz 180 deg; joints [-15.406, -58.924, 128.112, 163.575, 69.969, -84.234]
  MoveL 3860 to (0, 0, 58.6) mm, rotated rx 180 ry 0 rz 180 deg; joints [-13.245, -50.958, 111.986, 164.941, 61.869, -82.77]
  MoveL 3861 to (0, 0, 59) mm, rotated rx 180 ry 0 rz 180 deg; joints [-13.261, -50.954, 111.978, 164.923, 61.867, -82.761]
  MoveL 3862 to (-200, 0, 59) mm, rotated rx 180 ry 0 rz 180 deg; joints [-15.424, -58.919, 128.103, 163.555, 69.966, -84.226]
  MoveL 3863 to (-200, -0.6, 59) mm, rotated rx 180 ry 0 rz 180 deg; joints [-15.424, -58.959, 128.103, 163.551, 69.928, -84.214]
  MoveL 3864 to (0, -0.6, 59) mm, rotated rx 180 ry 0 rz 180 deg; joints [-13.261, -50.986, 111.977, 164.918, 61.835, -82.751]
  MoveL 3865 to (0, -1.2, 59) mm, rotated rx 180 ry 0 rz 180 deg; joints [-13.261, -51.018, 111.977, 164.913, 61.804, -82.741]
  MoveL 3866 to (-200, -1.2, 59) mm, rotated rx 180 ry 0 rz 180 deg; joints [-15.424, -58.998, 128.102, 163.547, 69.89, -84.202]
  MoveL 3867 to (-200, -1.8, 59) mm, rotated rx 180 ry 0 rz 180 deg; joints [-15.424, -59.037, 128.101, 163.543, 69.851, -84.19]
  MoveL 3868 to (0, -1.8, 59) mm, rotated rx 180 ry 0 rz 180 deg; joints [-13.261, -51.05, 111.976, 164.909, 61.772, -82.732]
  MoveL 3869 to (0, -2.4, 59) mm, rotated rx 180 ry 0 rz 180 deg; joints [-13.261, -51.082, 111.975, 164.904, 61.74, -82.722]
  MoveL 3870 to (-200, -2.4, 59) mm, rotated rx 180 ry 0 rz 180 deg; joints [-15.424, -59.077, 128.1, 163.539, 69.813, -84.178]
  MoveL 3871 to (-200, -3, 59) mm, rotated rx 180 ry 0 rz 180 deg; joints [-15.424, -59.116, 128.099, 163.535, 69.774, -84.166]
  MoveL 3872 to (0, -3, 59) mm, rotated rx 180 ry 0 rz 180 deg; joints [-13.261, -51.114, 111.974, 164.9, 61.708, -82.712]
  MoveL 3873 to (0, -3.6, 59) mm, rotated rx 180 ry 0 rz 180 deg; joints [-13.261, -51.146, 111.973, 164.895, 61.677, -82.702]
  MoveL 3874 to (-200, -3.6, 59) mm, rotated rx 180 ry 0 rz 180 deg; joints [-15.424, -59.155, 128.098, 163.53, 69.736, -84.154]
  MoveL 3875 to (-200, -4.2, 59) mm, rotated rx 180 ry 0 rz 180 deg; joints [-15.424, -59.194, 128.097, 163.526, 69.697, -84.141]
  MoveL 3876 to (0, -4.2, 59) mm, rotated rx 180 ry 0 rz 180 deg; joints [-13.261, -51.178, 111.973, 164.89, 61.645, -82.693]
  MoveL 3877 to (0, -4.8, 59) mm, rotated rx 180 ry 0 rz 180 deg; joints [-13.261, -51.21, 111.972, 164.886, 61.613, -82.683]
  MoveL 3878 to (-200, -4.8, 59) mm, rotated rx 180 ry 0 rz 180 deg; joints [-15.424, -59.234, 128.096, 163.522, 69.658, -84.129]
  MoveL 3879 to (-200, -5.4, 59) mm, rotated rx 180 ry 0 rz 180 deg; joints [-15.424, -59.273, 128.095, 163.518, 69.62, -84.117]
  MoveL 3880 to (0, -5.4, 59) mm, rotated rx 180 ry 0 rz 180 deg; joints [-13.261, -51.242, 111.971, 164.881, 61.582, -82.673]
  MoveL 3881 to (0, -6, 59) mm, rotated rx 180 ry 0 rz 180 deg; joints [-13.261, -51.274, 111.97, 164.877, 61.55, -82.664]
  MoveL 3882 to (-200, -6, 59) mm, rotated rx 180 ry 0 rz 180 deg; joints [-15.424, -59.312, 128.094, 163.514, 69.581, -84.105]
  MoveL 3883 to (-200, -6.6, 59) mm, rotated rx 180 ry 0 rz 180 deg; joints [-15.424, -59.351, 128.093, 163.509, 69.543, -84.093]
  MoveL 3884 to (0, -6.6, 59) mm, rotated rx 180 ry 0 rz 180 deg; joints [-13.261, -51.306, 111.969, 164.872, 61.518, -82.654]
  MoveL 3885 to (0, -7.2, 59) mm, rotated rx 180 ry 0 rz 180 deg; joints [-13.261, -51.338, 111.968, 164.867, 61.486, -82.644]
  MoveL 3886 to (-200, -7.2, 59) mm, rotated rx 180 ry 0 rz 180 deg; joints [-15.424, -59.39, 128.092, 163.505, 69.504, -84.081]
  MoveL 3887 to (-200, -7.8, 59) mm, rotated rx 180 ry 0 rz 180 deg; joints [-15.424, -59.43, 128.091, 163.501, 69.466, -84.068]
  MoveL 3888 to (0, -7.8, 59) mm, rotated rx 180 ry 0 rz 180 deg; joints [-13.261, -51.37, 111.967, 164.863, 61.454, -82.634]
  MoveL 3889 to (0, -8.4, 59) mm, rotated rx 180 ry 0 rz 180 deg; joints [-13.261, -51.402, 111.966, 164.858, 61.423, -82.624]
  MoveL 3890 to (-200, -8.4, 59) mm, rotated rx 180 ry 0 rz 180 deg; joints [-15.424, -59.469, 128.09, 163.496, 69.427, -84.056]
  MoveL 3891 to (-200, -9, 59) mm, rotated rx 180 ry 0 rz 180 deg; joints [-15.424, -59.508, 128.089, 163.492, 69.388, -84.044]
  MoveL 3892 to (0, -9, 59) mm, rotated rx 180 ry 0 rz 180 deg; joints [-13.261, -51.434, 111.965, 164.853, 61.391, -82.615]
  MoveL 3893 to (0, -9.6, 59) mm, rotated rx 180 ry 0 rz 180 deg; joints [-13.261, -51.466, 111.964, 164.848, 61.359, -82.605]
  MoveL 3894 to (-200, -9.6, 59) mm, rotated rx 180 ry 0 rz 180 deg; joints [-15.424, -59.547, 128.088, 163.488, 69.35, -84.032]
  MoveL 3895 to (-200, -10.2, 59) mm, rotated rx 180 ry 0 rz 180 deg; joints [-15.424, -59.586, 128.086, 163.484, 69.311, -84.019]
  MoveL 3896 to (0, -10.2, 59) mm, rotated rx 180 ry 0 rz 180 deg; joints [-13.261, -51.498, 111.963, 164.844, 61.327, -82.595]
  MoveL 3897 to (0, -10.8, 59) mm, rotated rx 180 ry 0 rz 180 deg; joints [-13.261, -51.529, 111.961, 164.839, 61.295, -82.585]
  MoveL 3898 to (-200, -10.8, 59) mm, rotated rx 180 ry 0 rz 180 deg; joints [-15.424, -59.625, 128.085, 163.479, 69.272, -84.007]
  MoveL 3899 to (-200, -11.4, 59) mm, rotated rx 180 ry 0 rz 180 deg; joints [-15.424, -59.664, 128.084, 163.475, 69.234, -83.995]
  MoveL 3900 to (0, -11.4, 59) mm, rotated rx 180 ry 0 rz 180 deg; joints [-13.261, -51.561, 111.96, 164.834, 61.263, -82.575]
  MoveL 3901 to (0, -12, 59) mm, rotated rx 180 ry 0 rz 180 deg; joints [-13.261, -51.593, 111.959, 164.83, 61.231, -82.565]
  MoveL 3902 to (-200, -12, 59) mm, rotated rx 180 ry 0 rz 180 deg; joints [-15.424, -59.703, 128.082, 163.47, 69.195, -83.983]
  MoveL 3903 to (-200, -12.6, 59) mm, rotated rx 180 ry 0 rz 180 deg; joints [-15.424, -59.742, 128.081, 163.466, 69.156, -83.97]
  MoveL 3904 to (0, -12.6, 59) mm, rotated rx 180 ry 0 rz 180 deg; joints [-13.261, -51.625, 111.958, 164.825, 61.199, -82.555]
  MoveL 3905 to (0, -13.2, 59) mm, rotated rx 180 ry 0 rz 180 deg; joints [-13.261, -51.657, 111.956, 164.82, 61.167, -82.546]
  MoveL 3906 to (-200, -13.2, 59) mm, rotated rx 180 ry 0 rz 180 deg; joints [-15.424, -59.781, 128.08, 163.462, 69.117, -83.958]
  MoveL 3907 to (-200, -13.8, 59) mm, rotated rx 180 ry 0 rz 180 deg; joints [-15.424, -59.82, 128.078, 163.457, 69.079, -83.946]
  MoveL 3908 to (0, -13.8, 59) mm, rotated rx 180 ry 0 rz 180 deg; joints [-13.261, -51.689, 111.955, 164.815, 61.135, -82.536]
  MoveL 3909 to (0, -14.4, 59) mm, rotated rx 180 ry 0 rz 180 deg; joints [-13.261, -51.72, 111.954, 164.81, 61.104, -82.526]
  MoveL 3910 to (-200, -14.4, 59) mm, rotated rx 180 ry 0 rz 180 deg; joints [-15.424, -59.859, 128.077, 163.453, 69.04, -83.933]
  MoveL 3911 to (-200, -15, 59) mm, rotated rx 180 ry 0 rz 180 deg; joints [-15.424, -59.898, 128.075, 163.448, 69.001, -83.921]
  MoveL 3912 to (0, -15, 59) mm, rotated rx 180 ry 0 rz 180 deg; joints [-13.261, -51.752, 111.952, 164.806, 61.072, -82.516]
  MoveL 3913 to (0, -15.6, 59) mm, rotated rx 180 ry 0 rz 180 deg; joints [-13.261, -51.784, 111.951, 164.801, 61.04, -82.506]
  MoveL 3914 to (-200, -15.6, 59) mm, rotated rx 180 ry 0 rz 180 deg; joints [-15.424, -59.937, 128.073, 163.444, 68.962, -83.909]
  MoveL 3915 to (-200, -16.2, 59) mm, rotated rx 180 ry 0 rz 180 deg; joints [-15.424, -59.976, 128.072, 163.44, 68.923, -83.896]
  MoveL 3916 to (0, -16.2, 59) mm, rotated rx 180 ry 0 rz 180 deg; joints [-13.261, -51.816, 111.95, 164.796, 61.008, -82.496]
  MoveL 3917 to (0, -16.8, 59) mm, rotated rx 180 ry 0 rz 180 deg; joints [-13.261, -51.847, 111.948, 164.791, 60.976, -82.486]
  MoveL 3918 to (-200, -16.8, 59) mm, rotated rx 180 ry 0 rz 180 deg; joints [-15.424, -60.015, 128.07, 163.435, 68.885, -83.884]
  MoveL 3919 to (-200, -17.4, 59) mm, rotated rx 180 ry 0 rz 180 deg; joints [-15.424, -60.054, 128.069, 163.431, 68.846, -83.871]
  MoveL 3920 to (0, -17.4, 59) mm, rotated rx 180 ry 0 rz 180 deg; joints [-13.261, -51.879, 111.947, 164.786, 60.944, -82.476]
  MoveL 3921 to (0, -18, 59) mm, rotated rx 180 ry 0 rz 180 deg; joints [-13.261, -51.911, 111.945, 164.782, 60.912, -82.466]
  MoveL 3922 to (-200, -18, 59) mm, rotated rx 180 ry 0 rz 180 deg; joints [-15.424, -60.092, 128.067, 163.426, 68.807, -83.859]
  MoveL 3923 to (-200, -18.6, 59) mm, rotated rx 180 ry 0 rz 180 deg; joints [-15.424, -60.131, 128.065, 163.422, 68.768, -83.847]
  MoveL 3924 to (0, -18.6, 59) mm, rotated rx 180 ry 0 rz 180 deg; joints [-13.261, -51.942, 111.944, 164.777, 60.879, -82.456]
  MoveL 3925 to (0, -19.2, 59) mm, rotated rx 180 ry 0 rz 180 deg; joints [-13.261, -51.974, 111.942, 164.772, 60.847, -82.446]
  MoveL 3926 to (-200, -19.2, 59) mm, rotated rx 180 ry 0 rz 180 deg; joints [-15.424, -60.17, 128.063, 163.417, 68.729, -83.834]
  MoveL 3927 to (-200, -19.8, 59) mm, rotated rx 180 ry 0 rz 180 deg; joints [-15.424, -60.209, 128.062, 163.413, 68.69, -83.822]
  MoveL 3928 to (0, -19.8, 59) mm, rotated rx 180 ry 0 rz 180 deg; joints [-13.261, -52.006, 111.94, 164.767, 60.815, -82.436]
  MoveL 3929 to (0, -20.4, 59) mm, rotated rx 180 ry 0 rz 180 deg; joints [-13.261, -52.037, 111.939, 164.762, 60.783, -82.426]
  MoveL 3930 to (-200, -20.4, 59) mm, rotated rx 180 ry 0 rz 180 deg; joints [-15.424, -60.248, 128.06, 163.408, 68.651, -83.809]
  MoveL 3931 to (-200, -21, 59) mm, rotated rx 180 ry 0 rz 180 deg; joints [-15.424, -60.286, 128.058, 163.404, 68.612, -83.797]
  MoveL 3932 to (0, -21, 59) mm, rotated rx 180 ry 0 rz 180 deg; joints [-13.261, -52.069, 111.937, 164.757, 60.751, -82.416]
  MoveL 3933 to (0, -21.6, 59) mm, rotated rx 180 ry 0 rz 180 deg; joints [-13.261, -52.1, 111.935, 164.752, 60.719, -82.406]
  MoveL 3934 to (-200, -21.6, 59) mm, rotated rx 180 ry 0 rz 180 deg; joints [-15.424, -60.325, 128.056, 163.399, 68.574, -83.784]
  MoveL 3935 to (-200, -22.2, 59) mm, rotated rx 180 ry 0 rz 180 deg; joints [-15.424, -60.364, 128.054, 163.395, 68.535, -83.772]
  MoveL 3936 to (0, -22.2, 59) mm, rotated rx 180 ry 0 rz 180 deg; joints [-13.261, -52.132, 111.934, 164.747, 60.687, -82.396]
  MoveL 3937 to (0, -22.8, 59) mm, rotated rx 180 ry 0 rz 180 deg; joints [-13.261, -52.163, 111.932, 164.742, 60.655, -82.386]
  MoveL 3938 to (-200, -22.8, 59) mm, rotated rx 180 ry 0 rz 180 deg; joints [-15.424, -60.402, 128.052, 163.39, 68.496, -83.76]
  MoveL 3939 to (-200, -23.4, 59) mm, rotated rx 180 ry 0 rz 180 deg; joints [-15.424, -60.441, 128.05, 163.385, 68.457, -83.747]
  MoveL 3940 to (0, -23.4, 59) mm, rotated rx 180 ry 0 rz 180 deg; joints [-13.261, -52.195, 111.93, 164.737, 60.623, -82.376]
  MoveL 3941 to (0, -24, 59) mm, rotated rx 180 ry 0 rz 180 deg; joints [-13.261, -52.227, 111.928, 164.733, 60.59, -82.366]
  MoveL 3942 to (-200, -24, 59) mm, rotated rx 180 ry 0 rz 180 deg; joints [-15.424, -60.48, 128.048, 163.381, 68.418, -83.734]
  MoveL 3943 to (-200, -24.6, 59) mm, rotated rx 180 ry 0 rz 180 deg; joints [-15.424, -60.518, 128.046, 163.376, 68.379, -83.722]
  MoveL 3944 to (0, -24.6, 59) mm, rotated rx 180 ry 0 rz 180 deg; joints [-13.261, -52.258, 111.926, 164.728, 60.558, -82.356]
  MoveL 3945 to (0, -25.2, 59) mm, rotated rx 180 ry 0 rz 180 deg; joints [-13.261, -52.29, 111.924, 164.723, 60.526, -82.346]
  MoveL 3946 to (-200, -25.2, 59) mm, rotated rx 180 ry 0 rz 180 deg; joints [-15.424, -60.557, 128.044, 163.372, 68.34, -83.709]
  MoveL 3947 to (-200, -25.8, 59) mm, rotated rx 180 ry 0 rz 180 deg; joints [-15.424, -60.596, 128.042, 163.367, 68.301, -83.697]
  MoveL 3948 to (0, -25.8, 59) mm, rotated rx 180 ry 0 rz 180 deg; joints [-13.261, -52.321, 111.923, 164.718, 60.494, -82.336]
  MoveL 3949 to (0, -26.4, 59) mm, rotated rx 180 ry 0 rz 180 deg; joints [-13.261, -52.352, 111.921, 164.713, 60.462, -82.325]
  MoveL 3950 to (-200, -26.4, 59) mm, rotated rx 180 ry 0 rz 180 deg; joints [-15.424, -60.634, 128.04, 163.362, 68.262, -83.684]
  MoveL 3951 to (-200, -27, 59) mm, rotated rx 180 ry 0 rz 180 deg; joints [-15.424, -60.673, 128.038, 163.358, 68.223, -83.672]
  MoveL 3952 to (0, -27, 59) mm, rotated rx 180 ry 0 rz 180 deg; joints [-13.261, -52.384, 111.919, 164.708, 60.429, -82.315]
  MoveL 3953 to (0, -27.6, 59) mm, rotated rx 180 ry 0 rz 180 deg; joints [-13.261, -52.415, 111.917, 164.703, 60.397, -82.305]
  MoveL 3954 to (-200, -27.6, 59) mm, rotated rx 180 ry 0 rz 180 deg; joints [-15.424, -60.711, 128.035, 163.353, 68.183, -83.659]
  MoveL 3955 to (-200, -28.2, 59) mm, rotated rx 180 ry 0 rz 180 deg; joints [-15.424, -60.75, 128.033, 163.348, 68.144, -83.647]
  MoveL 3956 to (0, -28.2, 59) mm, rotated rx 180 ry 0 rz 180 deg; joints [-13.261, -52.447, 111.915, 164.698, 60.365, -82.295]
  MoveL 3957 to (0, -28.8, 59) mm, rotated rx 180 ry 0 rz 180 deg; joints [-13.261, -52.478, 111.913, 164.693, 60.333, -82.285]
  MoveL 3958 to (-200, -28.8, 59) mm, rotated rx 180 ry 0 rz 180 deg; joints [-15.424, -60.788, 128.031, 163.344, 68.105, -83.634]
  MoveL 3959 to (-200, -29.4, 59) mm, rotated rx 180 ry 0 rz 180 deg; joints [-15.424, -60.827, 128.029, 163.339, 68.066, -83.621]
  MoveL 3960 to (0, -29.4, 59) mm, rotated rx 180 ry 0 rz 180 deg; joints [-13.261, -52.509, 111.91, 164.688, 60.3, -82.275]
  MoveL 3961 to (0, -30, 59) mm, rotated rx 180 ry 0 rz 180 deg; joints [-13.261, -52.541, 111.908, 164.683, 60.268, -82.264]
  MoveL 3962 to (-200, -30, 59) mm, rotated rx 180 ry 0 rz 180 deg; joints [-15.424, -60.865, 128.026, 163.334, 68.027, -83.609]
  MoveL 3963 to (-200, -30.6, 58.99) mm, rotated rx 177.54 ry 0 rz 180 deg; joints [-15.492, -61.865, 127.92, 163.128, 66.975, -85.691]
  MoveL 3964 to (0, -30.6, 58.99) mm, rotated rx 177.54 ry 0 rz 180 deg; joints [-13.321, -53.354, 111.811, 164.473, 59.399, -84.406]
  MoveL 3965 to (0, -31.2, 58.95) mm, rotated rx 175.09 ry 0 rz 180 deg; joints [-13.354, -54.163, 111.705, 164.287, 58.522, -86.554]
  MoveL 3966 to (-200, -31.2, 58.95) mm, rotated rx 175.09 ry 0 rz 180 deg; joints [-15.53, -62.861, 127.804, 162.946, 65.917, -87.776]
  MoveL 3967 to (-200, -31.8, 58.88) mm, rotated rx 172.63 ry 0 rz 180 deg; joints [-15.536, -63.852, 127.679, 162.789, 64.852, -89.868]
  MoveL 3968 to (0, -31.8, 58.88) mm, rotated rx 172.63 ry 0 rz 180 deg; joints [-13.359, -54.97, 111.592, 164.125, 57.638, -88.712]
  MoveL 3969 to (0, -32.39, 58.8) mm, rotated rx 170.18 ry 0 rz 180 deg; joints [-13.337, -55.77, 111.472, 163.988, 56.75, -90.88]
  MoveL 3970 to (-200, -32.39, 58.8) mm, rotated rx 170.18 ry 0 rz 180 deg; joints [-15.511, -64.835, 127.546, 162.657, 63.783, -91.967]
  MoveL 3971 to (-200, -32.98, 58.68) mm, rotated rx 167.72 ry 0 rz 180 deg; joints [-15.455, -65.809, 127.404, 162.551, 62.71, -94.077]
  MoveL 3972 to (0, -32.98, 58.68) mm, rotated rx 167.72 ry 0 rz 180 deg; joints [-13.288, -56.565, 111.345, 163.876, 55.857, -93.062]
  MoveL 3973 to (0, -33.56, 58.54) mm, rotated rx 165.27 ry 0 rz 180 deg; joints [-13.213, -57.35, 111.212, 163.79, 54.962, -95.257]
  MoveL 3974 to (-200, -33.56, 58.54) mm, rotated rx 165.27 ry 0 rz 180 deg; joints [-15.368, -66.772, 127.254, 162.472, 61.636, -96.2]
  MoveL 3975 to (-200, -34.14, 58.38) mm, rotated rx 162.81 ry 0 rz 180 deg; joints [-15.25, -67.722, 127.097, 162.421, 60.562, -98.339]
  MoveL 3976 to (0, -34.14, 58.38) mm, rotated rx 162.81 ry 0 rz 180 deg; joints [-13.11, -58.126, 111.072, 163.732, 54.065, -97.471]
  MoveL 3977 to (0, -34.71, 58.19) mm, rotated rx 160.36 ry 0 rz 180 deg; joints [-12.98, -58.891, 110.926, 163.703, 53.168, -99.703]
  MoveL 3978 to (-200, -34.71, 58.19) mm, rotated rx 160.36 ry 0 rz 180 deg; joints [-15.101, -68.658, 126.932, 162.399, 59.49, -100.495]
  MoveL 3979 to (-200, -35.27, 57.97) mm, rotated rx 157.9 ry 0 rz 180 deg; joints [-14.921, -69.578, 126.761, 162.408, 58.42, -102.672]
  MoveL 3980 to (0, -35.27, 57.97) mm, rotated rx 157.9 ry 0 rz 180 deg; joints [-12.823, -59.644, 110.774, 163.703, 52.273, -101.957]
  MoveL 3981 to (0, -35.82, 57.73) mm, rotated rx 155.44 ry 0 rz 180 deg; joints [-12.64, -60.383, 110.617, 163.735, 51.381, -104.235]
  MoveL 3982 to (-200, -35.82, 57.73) mm, rotated rx 155.44 ry 0 rz 180 deg; joints [-14.71, -70.481, 126.584, 162.448, 57.355, -104.873]
  MoveL 3983 to (-200, -36.36, 57.47) mm, rotated rx 152.99 ry 0 rz 180 deg; joints [-14.469, -71.365, 126.401, 162.522, 56.297, -107.1]
  MoveL 3984 to (0, -36.36, 57.47) mm, rotated rx 152.99 ry 0 rz 180 deg; joints [-12.431, -61.107, 110.456, 163.799, 50.492, -106.539]
  MoveL 3985 to (0, -36.89, 57.19) mm, rotated rx 150.53 ry 0 rz 180 deg; joints [-12.196, -61.816, 110.291, 163.897, 49.61, -108.871]
  MoveL 3986 to (-200, -36.89, 57.19) mm, rotated rx 150.53 ry 0 rz 180 deg; joints [-14.198, -72.229, 126.213, 162.63, 55.246, -109.356]
  MoveL 3987 to (-200, -37.4, 56.88) mm, rotated rx 148.08 ry 0 rz 180 deg; joints [-13.898, -73.071, 126.02, 162.775, 54.205, -111.644]
  MoveL 3988 to (0, -37.4, 56.88) mm, rotated rx 148.08 ry 0 rz 180 deg; joints [-11.934, -62.507, 110.121, 164.031, 48.735, -111.234]
  MoveL 3989 to (0, -37.91, 56.55) mm, rotated rx 145.62 ry 0 rz 180 deg; joints [-11.648, -63.18, 109.949, 164.202, 47.869, -113.63]
  MoveL 3990 to (-200, -37.91, 56.55) mm, rotated rx 145.62 ry 0 rz 180 deg; joints [-13.567, -73.89, 125.824, 162.959, 53.176, -113.967]
  MoveL 3991 to (-200, -38.39, 56.2) mm, rotated rx 143.17 ry 0 rz 180 deg; joints [-13.208, -74.685, 125.625, 163.183, 52.16, -116.329]
  MoveL 3992 to (0, -38.39, 56.2) mm, rotated rx 143.17 ry 0 rz 180 deg; joints [-11.336, -63.834, 109.774, 164.412, 47.013, -116.063]
  MoveL 3993 to (0, -38.87, 55.84) mm, rotated rx 140.71 ry 0 rz 180 deg; joints [-11, -64.468, 109.598, 164.662, 46.169, -118.534]
  MoveL 3994 to (-200, -38.87, 55.84) mm, rotated rx 140.71 ry 0 rz 180 deg; joints [-12.82, -75.455, 125.424, 163.449, 51.159, -118.731]
  MoveL 3995 to (-200, -39.32, 55.45) mm, rotated rx 138.26 ry 0 rz 180 deg; joints [-12.404, -76.198, 125.222, 163.759, 50.176, -121.176]
  MoveL 3996 to (0, -39.32, 55.45) mm, rotated rx 138.26 ry 0 rz 180 deg; joints [-10.64, -65.08, 109.42, 164.954, 45.34, -121.045]
  MoveL 3997 to (0, -39.76, 55.04) mm, rotated rx 135.8 ry 0 rz 180 deg; joints [-10.256, -65.67, 109.241, 165.291, 44.526, -123.599]
  MoveL 3998 to (-200, -39.76, 55.04) mm, rotated rx 135.8 ry 0 rz 180 deg; joints [-11.96, -76.913, 125.018, 164.115, 49.211, -123.669]
  MoveL 3999 to (-200, -40.18, 54.61) mm, rotated rx 133.34 ry 0 rz 180 deg; joints [-11.489, -77.6, 124.815, 164.52, 48.268, -126.21]
  MoveL 4000 to (0, -40.18, 54.61) mm, rotated rx 133.34 ry 0 rz 180 deg; joints [-9.85, -66.237, 109.063, 165.672, 43.73, -126.198]
  MoveL 4001 to (0, -40.58, 54.16) mm, rotated rx 130.89 ry 0 rz 180 deg; joints [-9.42, -66.78, 108.885, 166.101, 42.953, -128.845]
  MoveL 4002 to (-200, -40.58, 54.16) mm, rotated rx 130.89 ry 0 rz 180 deg; joints [-10.992, -78.258, 124.613, 164.975, 47.349, -128.804]
  MoveL 4003 to (-200, -40.97, 53.7) mm, rotated rx 128.43 ry 0 rz 180 deg; joints [-10.469, -78.885, 124.412, 165.482, 46.456, -131.451]
  MoveL 4004 to (0, -40.97, 53.7) mm, rotated rx 128.43 ry 0 rz 180 deg; joints [-8.97, -67.298, 108.709, 166.578, 42.199, -131.541]
  MoveL 4005 to (0, -41.33, 53.23) mm, rotated rx 125.98 ry 0 rz 180 deg; joints [-8.498, -67.791, 108.534, 167.106, 41.468, -134.288]
  MoveL 4006 to (-200, -41.33, 53.23) mm, rotated rx 125.98 ry 0 rz 180 deg; joints [-9.921, -79.482, 124.214, 166.043, 45.59, -134.156]
  MoveL 4007 to (-200, -41.67, 52.73) mm, rotated rx 123.52 ry 0 rz 180 deg; joints [-9.35, -80.046, 124.019, 166.66, 44.756, -136.919]
  MoveL 4008 to (0, -41.67, 52.73) mm, rotated rx 123.52 ry 0 rz 180 deg; joints [-8.006, -68.258, 108.362, 167.684, 40.763, -137.087]
  MoveL 4009 to (0, -41.99, 52.23) mm, rotated rx 121.07 ry 0 rz 180 deg; joints [-7.494, -68.699, 108.194, 168.314, 40.085, -139.941]
  MoveL 4010 to (-200, -41.99, 52.23) mm, rotated rx 121.07 ry 0 rz 180 deg; joints [-8.755, -80.577, 123.827, 167.333, 43.955, -139.742]
  MoveL 4011 to (-200, -42.29, 51.7) mm, rotated rx 118.61 ry 0 rz 180 deg; joints [-8.138, -81.075, 123.641, 168.063, 43.191, -142.626]
  MoveL 4012 to (0, -42.29, 51.7) mm, rotated rx 118.61 ry 0 rz 180 deg; joints [-6.964, -69.111, 108.029, 168.996, 39.439, -142.848]
  MoveL 4013 to (0, -42.57, 51.17) mm, rotated rx 116.16 ry 0 rz 180 deg; joints [-6.417, -69.496, 107.869, 169.731, 38.824, -145.81]
  MoveL 4014 to (-200, -42.57, 51.17) mm, rotated rx 116.16 ry 0 rz 180 deg; joints [-7.5, -81.539, 123.46, 168.852, 42.464, -145.573]
  MoveL 4015 to (-200, -42.82, 50.63) mm, rotated rx 113.7 ry 0 rz 180 deg; joints [-6.843, -81.968, 123.286, 169.699, 41.779, -148.58]
  MoveL 4016 to (0, -42.82, 50.63) mm, rotated rx 113.7 ry 0 rz 180 deg; joints [-5.853, -69.853, 107.715, 170.518, 38.244, -148.826]
  MoveL 4017 to (0, -43.05, 50.07) mm, rotated rx 111.25 ry 0 rz 180 deg; joints [-5.273, -70.18, 107.565, 171.357, 37.701, -151.897]
  MoveL 4018 to (-200, -43.05, 50.07) mm, rotated rx 111.25 ry 0 rz 180 deg; joints [-6.167, -82.363, 123.118, 170.603, 41.138, -151.65]
  MoveL 4019 to (-200, -43.25, 49.51) mm, rotated rx 108.79 ry 0 rz 180 deg; joints [-5.473, -82.722, 122.958, 171.562, 40.544, -154.778]
  MoveL 4020 to (0, -43.25, 49.51) mm, rotated rx 108.79 ry 0 rz 180 deg; joints [-4.679, -70.478, 107.423, 172.245, 37.198, -155.019]
  MoveL 4021 to (0, -43.44, 48.94) mm, rotated rx 106.33 ry 0 rz 180 deg; joints [-4.072, -70.747, 107.287, 173.182, 36.735, -158.192]
  MoveL 4022 to (-200, -43.44, 48.94) mm, rotated rx 106.33 ry 0 rz 180 deg; joints [-4.764, -83.044, 122.806, 172.576, 39.998, -157.966]
  MoveL 4023 to (-200, -43.59, 48.36) mm, rotated rx 103.88 ry 0 rz 180 deg; joints [-4.04, -83.331, 122.662, 173.642, 39.505, -161.208]
  MoveL 4024 to (0, -43.59, 48.36) mm, rotated rx 103.88 ry 0 rz 180 deg; joints [-3.452, -70.985, 107.159, 174.164, 36.315, -161.414]
  MoveL 4025 to (0, -43.72, 47.77) mm, rotated rx 101.42 ry 0 rz 180 deg; joints [-2.822, -71.194, 107.038, 175.188, 35.94, -164.678]
  MoveL 4026 to (-200, -43.72, 47.77) mm, rotated rx 101.42 ry 0 rz 180 deg; joints [-3.303, -83.581, 122.529, 174.754, 39.065, -164.5]
  MoveL 4027 to (-200, -43.83, 47.18) mm, rotated rx 98.97 ry 0 rz 180 deg; joints [-2.555, -83.794, 122.404, 175.911, 38.682, -167.839]
  MoveL 4028 to (0, -43.83, 47.18) mm, rotated rx 98.97 ry 0 rz 180 deg; joints [-2.183, -71.371, 106.926, 176.25, 35.613, -167.983]
  MoveL 4029 to (0, -43.91, 46.59) mm, rotated rx 96.51 ry 0 rz 180 deg; joints [-1.535, -71.518, 106.822, 177.346, 35.333, -171.322]
  MoveL 4030 to (-200, -43.91, 46.59) mm, rotated rx 96.51 ry 0 rz 180 deg; joints [-1.797, -83.97, 122.291, 177.104, 38.357, -171.217]
  MoveL 4031 to (-200, -43.97, 45.99) mm, rotated rx 94.06 ry 0 rz 180 deg; joints [-1.03, -84.108, 122.188, 178.331, 38.091, -174.63]
  MoveL 4032 to (0, -43.97, 45.99) mm, rotated rx 94.06 ry 0 rz 180 deg; joints [-0.88, -71.634, 106.728, 178.47, 35.103, -174.692]
  MoveL 4033 to (0, -43.99, 45.39) mm, rotated rx 91.6 ry 0 rz 180 deg; joints [-0.219, -71.719, 106.643, 179.617, 34.924, -178.085]
  MoveL 4034 to (-200, -43.99, 45.39) mm, rotated rx 91.6 ry 0 rz 180 deg; joints [-0.257, -84.21, 122.096, 179.582, 37.887, -178.069]
  MoveL 4035 to (-200, -44, 44.79) mm, rotated rx 90 ry 0 rz 180 deg; joints [0.26, -84.255, 122.042, -179.575, 37.787, 179.664]
  MoveL 4036 to (0, -44, 44.79) mm, rotated rx 90 ry 0 rz 180 deg; joints [0.222, -71.757, 106.592, -179.611, 34.836, 179.681]
  MoveL 4037 to (0, -44, 44.19) mm, rotated rx 90 ry 0 rz 180 deg; joints [0.247, -71.757, 106.592, -179.567, 34.836, 179.645]
  MoveL 4038 to (-200, -44, 44.19) mm, rotated rx 90 ry 0 rz 180 deg; joints [0.29, -84.255, 122.041, -179.527, 37.787, 179.627]
  MoveL 4039 to (-200, -44, 43.59) mm, rotated rx 90 ry 0 rz 180 deg; joints [0.319, -84.255, 122.041, -179.48, 37.787, 179.589]
  MoveL 4040 to (0, -44, 43.59) mm, rotated rx 90 ry 0 rz 180 deg; joints [0.272, -71.757, 106.592, -179.523, 34.836, 179.609]
  MoveL 4041 to (0, -44, 42.99) mm, rotated rx 90 ry 0 rz 180 deg; joints [0.297, -71.757, 106.591, -179.479, 34.836, 179.573]
  MoveL 4042 to (-200, -44, 42.99) mm, rotated rx 90 ry 0 rz 180 deg; joints [0.348, -84.255, 122.041, -179.432, 37.787, 179.551]
  MoveL 4043 to (-200, -44, 42.39) mm, rotated rx 90 ry 0 rz 180 deg; joints [0.378, -84.255, 122.041, -179.384, 37.788, 179.513]
  MoveL 4044 to (0, -44, 42.39) mm, rotated rx 90 ry 0 rz 180 deg; joints [0.322, -71.757, 106.591, -179.435, 34.836, 179.537]
  MoveL 4045 to (0, -44, 41.79) mm, rotated rx 90 ry 0 rz 180 deg; joints [0.348, -71.756, 106.591, -179.392, 34.836, 179.501]
  MoveL 4046 to (-200, -44, 41.79) mm, rotated rx 90 ry 0 rz 180 deg; joints [0.407, -84.254, 122.04, -179.336, 37.788, 179.475]
  MoveL 4047 to (-200, -44, 41.19) mm, rotated rx 90 ry 0 rz 180 deg; joints [0.436, -84.254, 122.04, -179.288, 37.788, 179.437]
  MoveL 4048 to (0, -44, 41.19) mm, rotated rx 90 ry 0 rz 180 deg; joints [0.373, -71.756, 106.591, -179.348, 34.836, 179.465]
  MoveL 4049 to (0, -44, 40.59) mm, rotated rx 90 ry 0 rz 180 deg; joints [0.398, -71.756, 106.59, -179.304, 34.836, 179.429]
  MoveL 4050 to (-200, -44, 40.59) mm, rotated rx 90 ry 0 rz 180 deg; joints [0.466, -84.254, 122.04, -179.24, 37.788, 179.4]
  MoveL 4051 to (-200, -44, 39.99) mm, rotated rx 90 ry 0 rz 180 deg; joints [0.495, -84.253, 122.039, -179.192, 37.789, 179.362]
  MoveL 4052 to (0, -44, 39.99) mm, rotated rx 90 ry 0 rz 180 deg; joints [0.423, -71.756, 106.59, -179.26, 34.837, 179.393]
  MoveL 4053 to (0, -44, 39.39) mm, rotated rx 90 ry 0 rz 180 deg; joints [0.448, -71.755, 106.59, -179.216, 34.837, 179.357]
  MoveL 4054 to (-200, -44, 39.39) mm, rotated rx 90 ry 0 rz 180 deg; joints [0.524, -84.253, 122.039, -179.145, 37.789, 179.324]
  MoveL 4055 to (-200, -44, 38.79) mm, rotated rx 90 ry 0 rz 180 deg; joints [0.554, -84.253, 122.038, -179.097, 37.789, 179.286]
  MoveL 4056 to (0, -44, 38.79) mm, rotated rx 90 ry 0 rz 180 deg; joints [0.473, -71.755, 106.589, -179.172, 34.837, 179.321]
  MoveL 4057 to (0, -44, 38.19) mm, rotated rx 90 ry 0 rz 180 deg; joints [0.498, -71.755, 106.589, -179.128, 34.837, 179.285]
  MoveL 4058 to (-200, -44, 38.19) mm, rotated rx 90 ry 0 rz 180 deg; joints [0.583, -84.252, 122.038, -179.049, 37.79, 179.248]
  MoveL 4059 to (-200, -44, 37.59) mm, rotated rx 90 ry 0 rz 180 deg; joints [0.612, -84.252, 122.038, -179.001, 37.79, 179.21]
  MoveL 4060 to (0, -44, 37.59) mm, rotated rx 90 ry 0 rz 180 deg; joints [0.523, -71.754, 106.588, -179.085, 34.837, 179.249]
  MoveL 4061 to (0, -44, 36.99) mm, rotated rx 90 ry 0 rz 180 deg; joints [0.548, -71.754, 106.588, -179.041, 34.838, 179.213]
  MoveL 4062 to (-200, -44, 36.99) mm, rotated rx 90 ry 0 rz 180 deg; joints [0.641, -84.252, 122.037, -178.953, 37.79, 179.173]
  MoveL 4063 to (-200, -44, 36.39) mm, rotated rx 90 ry 0 rz 180 deg; joints [0.671, -84.251, 122.037, -178.905, 37.791, 179.135]
  MoveL 4064 to (0, -44, 36.39) mm, rotated rx 90 ry 0 rz 180 deg; joints [0.573, -71.754, 106.587, -178.997, 34.838, 179.177]
  MoveL 4065 to (0, -44, 35.79) mm, rotated rx 90 ry 0 rz 180 deg; joints [0.598, -71.753, 106.587, -178.953, 34.838, 179.141]
  MoveL 4066 to (-200, -44, 35.79) mm, rotated rx 90 ry 0 rz 180 deg; joints [0.7, -84.251, 122.036, -178.857, 37.791, 179.097]
  MoveL 4067 to (-200, -44, 35.19) mm, rotated rx 90 ry 0 rz 180 deg; joints [0.729, -84.25, 122.036, -178.81, 37.791, 179.059]
  MoveL 4068 to (0, -44, 35.19) mm, rotated rx 90 ry 0 rz 180 deg; joints [0.623, -71.753, 106.586, -178.909, 34.838, 179.105]
  MoveL 4069 to (0, -44, 34.59) mm, rotated rx 90 ry 0 rz 180 deg; joints [0.648, -71.752, 106.586, -178.865, 34.838, 179.069]
  MoveL 4070 to (-200, -44, 34.59) mm, rotated rx 90 ry 0 rz 180 deg; joints [0.759, -84.25, 122.035, -178.762, 37.792, 179.021]
  MoveL 4071 to (-200, -44, 33.99) mm, rotated rx 90 ry 0 rz 180 deg; joints [0.788, -84.249, 122.034, -178.714, 37.792, 178.984]
  MoveL 4072 to (0, -44, 33.99) mm, rotated rx 90 ry 0 rz 180 deg; joints [0.673, -71.752, 106.585, -178.821, 34.839, 179.033]
  MoveL 4073 to (0, -44, 33.39) mm, rotated rx 90 ry 0 rz 180 deg; joints [0.698, -71.752, 106.585, -178.778, 34.839, 178.997]
  MoveL 4074 to (-200, -44, 33.39) mm, rotated rx 90 ry 0 rz 180 deg; joints [0.817, -84.249, 122.034, -178.666, 37.793, 178.946]
  MoveL 4075 to (-200, -44, 32.79) mm, rotated rx 90 ry 0 rz 180 deg; joints [0.847, -84.248, 122.033, -178.618, 37.793, 178.908]
  MoveL 4076 to (0, -44, 32.79) mm, rotated rx 90 ry 0 rz 180 deg; joints [0.723, -71.751, 106.584, -178.734, 34.839, 178.961]
  MoveL 4077 to (0, -44, 32.19) mm, rotated rx 90 ry 0 rz 180 deg; joints [0.748, -71.751, 106.583, -178.69, 34.84, 178.925]
  MoveL 4078 to (-200, -44, 32.19) mm, rotated rx 90 ry 0 rz 180 deg; joints [0.876, -84.247, 122.033, -178.57, 37.794, 178.87]
  MoveL 4079 to (-200, -44, 31.59) mm, rotated rx 90 ry 0 rz 180 deg; joints [0.905, -84.247, 122.032, -178.522, 37.794, 178.832]
  MoveL 4080 to (0, -44, 31.59) mm, rotated rx 90 ry 0 rz 180 deg; joints [0.773, -71.75, 106.583, -178.646, 34.84, 178.889]
  MoveL 4081 to (0, -44, 30.99) mm, rotated rx 90 ry 0 rz 180 deg; joints [0.799, -71.75, 106.582, -178.602, 34.84, 178.853]
  MoveL 4082 to (-200, -44, 30.99) mm, rotated rx 90 ry 0 rz 180 deg; joints [0.935, -84.246, 122.031, -178.475, 37.795, 178.794]
  MoveL 4083 to (-200, -44, 30.39) mm, rotated rx 90 ry 0 rz 180 deg; joints [0.964, -84.246, 122.031, -178.427, 37.795, 178.757]
  MoveL 4084 to (0, -44, 30.39) mm, rotated rx 90 ry 0 rz 180 deg; joints [0.824, -71.749, 106.581, -178.558, 34.841, 178.817]
  MoveL 4085 to (0, -44, 29.79) mm, rotated rx 90 ry 0 rz 180 deg; joints [0.849, -71.749, 106.58, -178.514, 34.841, 178.781]
  MoveL 4086 to (-200, -44, 29.79) mm, rotated rx 90 ry 0 rz 180 deg; joints [0.993, -84.245, 122.03, -178.379, 37.796, 178.719]
  MoveL 4087 to (-200, -44, 29.19) mm, rotated rx 90 ry 0 rz 180 deg; joints [1.023, -84.244, 122.029, -178.331, 37.797, 178.681]
  MoveL 4088 to (0, -44, 29.19) mm, rotated rx 90 ry 0 rz 180 deg; joints [0.874, -71.748, 106.58, -178.471, 34.841, 178.745]
  MoveL 4089 to (0, -44, 28.59) mm, rotated rx 90 ry 0 rz 180 deg; joints [0.899, -71.747, 106.579, -178.427, 34.842, 178.709]
  MoveL 4090 to (-200, -44, 28.59) mm, rotated rx 90 ry 0 rz 180 deg; joints [1.052, -84.244, 122.028, -178.283, 37.797, 178.643]
  MoveL 4091 to (-200, -44, 27.99) mm, rotated rx 90 ry 0 rz 180 deg; joints [1.081, -84.243, 122.027, -178.235, 37.798, 178.605]
  MoveL 4092 to (0, -44, 27.99) mm, rotated rx 90 ry 0 rz 180 deg; joints [0.924, -71.747, 106.578, -178.383, 34.842, 178.673]
  MoveL 4093 to (0, -44, 27.39) mm, rotated rx 90 ry 0 rz 180 deg; joints [0.949, -71.746, 106.577, -178.339, 34.842, 178.637]
  MoveL 4094 to (-200, -44, 27.39) mm, rotated rx 90 ry 0 rz 180 deg; joints [1.111, -84.242, 122.027, -178.188, 37.798, 178.568]
  MoveL 4095 to (-200, -44, 26.79) mm, rotated rx 90 ry 0 rz 180 deg; joints [1.14, -84.241, 122.026, -178.14, 37.799, 178.53]
  MoveL 4096 to (0, -44, 26.79) mm, rotated rx 90 ry 0 rz 180 deg; joints [0.974, -71.746, 106.576, -178.295, 34.843, 178.601]
  MoveL 4097 to (0, -44, 26.19) mm, rotated rx 90 ry 0 rz 180 deg; joints [0.999, -71.745, 106.576, -178.251, 34.843, 178.565]
  MoveL 4098 to (-200, -44, 26.19) mm, rotated rx 90 ry 0 rz 180 deg; joints [1.169, -84.241, 122.025, -178.092, 37.8, 178.492]
  MoveL 4099 to (-200, -44, 25.59) mm, rotated rx 90 ry 0 rz 180 deg; joints [1.199, -84.24, 122.024, -178.044, 37.8, 178.454]
  MoveL 4100 to (0, -44, 25.59) mm, rotated rx 90 ry 0 rz 180 deg; joints [1.024, -71.744, 106.575, -178.208, 34.844, 178.529]
  MoveL 4101 to (0, -44, 24.99) mm, rotated rx 90 ry 0 rz 180 deg; joints [1.049, -71.744, 106.574, -178.164, 34.844, 178.493]
  MoveL 4102 to (-200, -44, 24.99) mm, rotated rx 90 ry 0 rz 180 deg; joints [1.228, -84.239, 122.023, -177.996, 37.801, 178.416]
  MoveL 4103 to (-200, -44, 24.39) mm, rotated rx 90 ry 0 rz 180 deg; joints [1.257, -84.238, 122.022, -177.948, 37.802, 178.379]
  MoveL 4104 to (0, -44, 24.39) mm, rotated rx 90 ry 0 rz 180 deg; joints [1.074, -71.743, 106.573, -178.12, 34.844, 178.457]
  MoveL 4105 to (0, -44, 23.79) mm, rotated rx 90 ry 0 rz 180 deg; joints [1.099, -71.742, 106.572, -178.076, 34.845, 178.421]
  MoveL 4106 to (-200, -44, 23.79) mm, rotated rx 90 ry 0 rz 180 deg; joints [1.287, -84.237, 122.021, -177.901, 37.803, 178.341]
  MoveL 4107 to (-200, -44, 23.19) mm, rotated rx 90 ry 0 rz 180 deg; joints [1.316, -84.236, 122.02, -177.853, 37.803, 178.303]
  MoveL 4108 to (0, -44, 23.19) mm, rotated rx 90 ry 0 rz 180 deg; joints [1.124, -71.742, 106.571, -178.032, 34.845, 178.385]
  MoveL 4109 to (0, -44, 22.59) mm, rotated rx 90 ry 0 rz 180 deg; joints [1.149, -71.741, 106.57, -177.988, 34.846, 178.349]
  MoveL 4110 to (-200, -44, 22.59) mm, rotated rx 90 ry 0 rz 180 deg; joints [1.345, -84.235, 122.019, -177.805, 37.804, 178.265]
  MoveL 4111 to (-200, -44, 21.99) mm, rotated rx 90 ry 0 rz 180 deg; joints [1.375, -84.235, 122.018, -177.757, 37.805, 178.228]
  MoveL 4112 to (0, -44, 21.99) mm, rotated rx 90 ry 0 rz 180 deg; joints [1.174, -71.74, 106.569, -177.945, 34.846, 178.313]
  MoveL 4113 to (0, -44, 21.39) mm, rotated rx 90 ry 0 rz 180 deg; joints [1.199, -71.739, 106.568, -177.901, 34.847, 178.277]
  MoveL 4114 to (-200, -44, 21.39) mm, rotated rx 90 ry 0 rz 180 deg; joints [1.404, -84.234, 122.017, -177.709, 37.806, 178.19]
  MoveL 4115 to (-200, -44, 20.79) mm, rotated rx 90 ry 0 rz 180 deg; joints [1.433, -84.233, 122.016, -177.662, 37.807, 178.152]
  MoveL 4116 to (0, -44, 20.79) mm, rotated rx 90 ry 0 rz 180 deg; joints [1.224, -71.739, 106.567, -177.857, 34.847, 178.241]
  MoveL 4117 to (0, -44, 20.19) mm, rotated rx 90 ry 0 rz 180 deg; joints [1.249, -71.738, 106.566, -177.813, 34.848, 178.205]
  MoveL 4118 to (-200, -44, 20.19) mm, rotated rx 90 ry 0 rz 180 deg; joints [1.463, -84.232, 122.015, -177.614, 37.807, 178.114]
  MoveL 4119 to (-200, -44, 19.59) mm, rotated rx 90 ry 0 rz 180 deg; joints [1.492, -84.231, 122.014, -177.566, 37.808, 178.076]
  MoveL 4120 to (0, -44, 19.59) mm, rotated rx 90 ry 0 rz 180 deg; joints [1.274, -71.737, 106.565, -177.769, 34.848, 178.169]
  MoveL 4121 to (0, -44, 18.99) mm, rotated rx 90 ry 0 rz 180 deg; joints [1.299, -71.736, 106.564, -177.725, 34.849, 178.133]
  MoveL 4122 to (-200, -44, 18.99) mm, rotated rx 90 ry 0 rz 180 deg; joints [1.521, -84.23, 122.013, -177.518, 37.809, 178.039]
  MoveL 4123 to (-200, -44, 18.39) mm, rotated rx 90 ry 0 rz 180 deg; joints [1.55, -84.229, 122.012, -177.47, 37.81, 178.001]
  MoveL 4124 to (0, -44, 18.39) mm, rotated rx 90 ry 0 rz 180 deg; joints [1.325, -71.735, 106.562, -177.682, 34.849, 178.097]
  MoveL 4125 to (0, -44, 17.79) mm, rotated rx 90 ry 0 rz 180 deg; joints [1.35, -71.734, 106.561, -177.638, 34.85, 178.061]
  MoveL 4126 to (-200, -44, 17.79) mm, rotated rx 90 ry 0 rz 180 deg; joints [1.58, -84.228, 122.01, -177.423, 37.811, 177.963]
  MoveL 4127 to (-200, -44, 17.19) mm, rotated rx 90 ry 0 rz 180 deg; joints [1.609, -84.226, 122.009, -177.375, 37.812, 177.925]
  MoveL 4128 to (0, -44, 17.19) mm, rotated rx 90 ry 0 rz 180 deg; joints [1.375, -71.734, 106.56, -177.594, 34.85, 178.025]
  MoveL 4129 to (0, -44, 16.59) mm, rotated rx 90 ry 0 rz 180 deg; joints [1.4, -71.733, 106.559, -177.55, 34.851, 177.989]
  MoveL 4130 to (-200, -44, 16.59) mm, rotated rx 90 ry 0 rz 180 deg; joints [1.638, -84.225, 122.008, -177.327, 37.813, 177.888]
  MoveL 4131 to (-200, -44, 15.99) mm, rotated rx 90 ry 0 rz 180 deg; joints [1.668, -84.224, 122.007, -177.279, 37.814, 177.85]
  MoveL 4132 to (0, -44, 15.99) mm, rotated rx 90 ry 0 rz 180 deg; joints [1.425, -71.732, 106.558, -177.506, 34.851, 177.953]
  MoveL 4133 to (0, -44, 15.39) mm, rotated rx 90 ry 0 rz 180 deg; joints [1.45, -71.731, 106.556, -177.463, 34.852, 177.917]
  MoveL 4134 to (-200, -44, 15.39) mm, rotated rx 90 ry 0 rz 180 deg; joints [1.697, -84.223, 122.006, -177.231, 37.815, 177.812]
  MoveL 4135 to (-200, -44, 14.79) mm, rotated rx 89.14 ry 0 rz 180 deg; joints [1.987, -84.231, 121.968, -176.755, 37.781, 176.579]
  MoveL 4136 to (0, -44, 14.79) mm, rotated rx 89.14 ry 0 rz 180 deg; joints [1.698, -71.738, 106.52, -177.026, 34.819, 176.703]
  MoveL 4137 to (0, -43.98, 14.19) mm, rotated rx 86.69 ry 0 rz 180 deg; joints [2.364, -71.739, 106.426, -175.85, 34.757, 173.279]
  MoveL 4138 to (-200, -43.98, 14.19) mm, rotated rx 86.69 ry 0 rz 180 deg; joints [2.767, -84.232, 121.869, -175.475, 37.724, 173.108]
  MoveL 4139 to (-200, -43.93, 13.59) mm, rotated rx 84.23 ry 0 rz 180 deg; joints [3.548, -84.194, 121.782, -174.196, 37.73, 169.637]
  MoveL 4140 to (0, -43.93, 13.59) mm, rotated rx 84.23 ry 0 rz 180 deg; joints [3.032, -71.709, 106.341, -174.675, 34.748, 169.855]
  MoveL 4141 to (0, -43.86, 13) mm, rotated rx 81.78 ry 0 rz 180 deg; joints [3.699, -71.648, 106.266, -173.507, 34.79, 166.439]
  MoveL 4142 to (-200, -43.86, 13) mm, rotated rx 81.78 ry 0 rz 180 deg; joints [4.328, -84.12, 121.707, -172.927, 37.799, 166.179]
  MoveL 4143 to (-200, -43.76, 12.41) mm, rotated rx 79.32 ry 0 rz 180 deg; joints [5.106, -84.009, 121.644, -171.675, 37.929, 162.739]
  MoveL 4144 to (0, -43.76, 12.41) mm, rotated rx 79.32 ry 0 rz 180 deg; joints [4.365, -71.557, 106.201, -172.353, 34.885, 163.038]
  MoveL 4145 to (0, -43.63, 11.82) mm, rotated rx 76.87 ry 0 rz 180 deg; joints [5.027, -71.434, 106.147, -171.219, 35.03, 159.659]
  MoveL 4146 to (-200, -43.63, 11.82) mm, rotated rx 76.87 ry 0 rz 180 deg; joints [5.879, -83.861, 121.593, -170.448, 38.119, 159.327]
  MoveL 4147 to (-200, -43.48, 11.24) mm, rotated rx 74.41 ry 0 rz 180 deg; joints [6.647, -83.677, 121.553, -169.253, 38.369, 155.948]
  MoveL 4148 to (0, -43.48, 11.24) mm, rotated rx 74.41 ry 0 rz 180 deg; joints [5.685, -71.282, 106.103, -170.111, 35.225, 156.307]
  MoveL 4149 to (0, -43.31, 10.66) mm, rotated rx 71.96 ry 0 rz 180 deg; joints [6.337, -71.099, 106.07, -169.035, 35.468, 152.99]
  MoveL 4150 to (-200, -43.31, 10.66) mm, rotated rx 71.96 ry 0 rz 180 deg; joints [7.407, -83.458, 121.526, -168.095, 38.675, 152.61]
  MoveL 4151 to (-200, -43.11, 10.1) mm, rotated rx 69.5 ry 0 rz 180 deg; joints [8.158, -83.202, 121.51, -166.979, 39.036, 149.318]
  MoveL 4152 to (0, -43.11, 10.1) mm, rotated rx 69.5 ry 0 rz 180 deg; joints [6.981, -70.887, 106.046, -167.995, 35.758, 149.71]
  MoveL 4153 to (0, -42.89, 9.54) mm, rotated rx 67.05 ry 0 rz 180 deg; joints [7.617, -70.646, 106.033, -166.996, 36.093, 146.474]
  MoveL 4154 to (-200, -42.89, 9.54) mm, rotated rx 67.05 ry 0 rz 180 deg; joints [8.898, -82.912, 121.506, -165.911, 39.45, 146.077]
  MoveL 4155 to (-200, -42.65, 8.99) mm, rotated rx 64.59 ry 0 rz 180 deg; joints [9.626, -82.587, 121.513, -164.894, 39.914, 142.893]
  MoveL 4156 to (0, -42.65, 8.99) mm, rotated rx 64.59 ry 0 rz 180 deg; joints [8.244, -70.376, 106.029, -166.042, 36.471, 143.287]
  MoveL 4157 to (0, -42.38, 8.46) mm, rotated rx 62.13 ry 0 rz 180 deg; joints [8.859, -70.077, 106.036, -165.134, 36.89, 140.148]
  MoveL 4158 to (-200, -42.38, 8.46) mm, rotated rx 62.13 ry 0 rz 180 deg; joints [10.341, -82.229, 121.531, -163.93, 40.426, 139.765]
  MoveL 4159 to (-200, -42.09, 7.93) mm, rotated rx 59.68 ry 0 rz 180 deg; joints [11.04, -81.837, 121.56, -163.023, 40.982, 136.701]
  MoveL 4160 to (0, -42.09, 7.93) mm, rotated rx 59.68 ry 0 rz 180 deg; joints [9.462, -69.751, 106.052, -164.277, 37.348, 137.064]
  MoveL 4161 to (0, -41.77, 7.42) mm, rotated rx 57.22 ry 0 rz 180 deg; joints [10.052, -69.398, 106.076, -163.471, 37.844, 134.034]
  MoveL 4162 to (-200, -41.77, 7.42) mm, rotated rx 57.22 ry 0 rz 180 deg; joints [11.723, -81.412, 121.599, -162.173, 41.581, 133.697]
  MoveL 4163 to (-200, -41.44, 6.92) mm, rotated rx 54.77 ry 0 rz 180 deg; joints [12.389, -80.956, 121.648, -161.381, 42.22, 130.758]
  MoveL 4164 to (0, -41.44, 6.92) mm, rotated rx 54.77 ry 0 rz 180 deg; joints [10.627, -69.017, 106.11, -162.718, 38.374, 131.061]
  MoveL 4165 to (0, -41.08, 6.44) mm, rotated rx 52.31 ry 0 rz 180 deg; joints [11.188, -68.611, 106.153, -162.017, 38.937, 128.142]
  MoveL 4166 to (-200, -41.08, 6.44) mm, rotated rx 52.31 ry 0 rz 180 deg; joints [13.036, -80.468, 121.706, -160.647, 42.895, 127.882]
  MoveL 4167 to (-200, -40.7, 5.97) mm, rotated rx 49.86 ry 0 rz 180 deg; joints [13.663, -79.95, 121.773, -159.97, 43.605, 125.069]
  MoveL 4168 to (0, -40.7, 5.97) mm, rotated rx 49.86 ry 0 rz 180 deg; joints [11.731, -68.179, 106.203, -161.37, 39.529, 125.282]
  MoveL 4169 to (0, -40.31, 5.52) mm, rotated rx 47.4 ry 0 rz 180 deg; joints [12.258, -67.722, 106.261, -160.776, 40.151, 122.476]
  MoveL 4170 to (-200, -40.31, 5.52) mm, rotated rx 47.4 ry 0 rz 180 deg; joints [14.27, -79.402, 121.849, -159.351, 44.346, 122.318]
  MoveL 4171 to (-200, -39.89, 5.09) mm, rotated rx 44.95 ry 0 rz 180 deg; joints [14.855, -78.825, 121.933, -158.787, 45.116, 119.629]
  MoveL 4172 to (0, -39.89, 5.09) mm, rotated rx 44.95 ry 0 rz 180 deg; joints [12.766, -67.241, 106.327, -160.233, 40.798, 119.727]
  MoveL 4173 to (0, -39.46, 4.68) mm, rotated rx 42.49 ry 0 rz 180 deg; joints [13.256, -66.737, 106.399, -159.742, 41.469, 117.031]
  MoveL 4174 to (-200, -39.46, 4.68) mm, rotated rx 42.49 ry 0 rz 180 deg; joints [15.418, -78.22, 122.024, -158.277, 45.914, 116.997]
  MoveL 4175 to (-200, -39.01, 4.28) mm, rotated rx 40.03 ry 0 rz 180 deg; joints [15.956, -77.587, 122.122, -157.82, 46.736, 114.424]
  MoveL 4176 to (0, -39.01, 4.28) mm, rotated rx 40.03 ry 0 rz 180 deg; joints [13.725, -66.21, 106.478, -159.3, 42.163, 114.388]
  MoveL 4177 to (0, -38.54, 3.9) mm, rotated rx 37.58 ry 0 rz 180 deg; joints [14.175, -65.661, 106.562, -158.906, 42.877, 111.794]
  MoveL 4178 to (-200, -38.54, 3.9) mm, rotated rx 37.58 ry 0 rz 180 deg; joints [16.472, -76.928, 122.226, -157.413, 47.58, 111.904]
  MoveL 4179 to (-200, -38.05, 3.55) mm, rotated rx 35.12 ry 0 rz 180 deg; joints [16.962, -76.244, 122.336, -157.055, 48.445, 109.438]
  MoveL 4180 to (0, -38.05, 3.55) mm, rotated rx 35.12 ry 0 rz 180 deg; joints [14.603, -65.091, 106.652, -158.559, 43.608, 109.251]
  MoveL 4181 to (0, -37.56, 3.21) mm, rotated rx 32.67 ry 0 rz 180 deg; joints [15.01, -64.5, 106.748, -158.257, 44.357, 106.753]
  MoveL 4182 to (-200, -37.56, 3.21) mm, rotated rx 32.67 ry 0 rz 180 deg; joints [17.427, -75.536, 122.451, -156.743, 49.328, 107.02]
  MoveL 4183 to (-200, -37.05, 2.9) mm, rotated rx 30.21 ry 0 rz 180 deg; joints [17.866, -74.803, 122.57, -156.475, 50.228, 104.649]
  MoveL 4184 to (0, -37.05, 2.9) mm, rotated rx 30.21 ry 0 rz 180 deg; joints [15.394, -63.891, 106.847, -157.999, 45.121, 104.299]
  MoveL 4185 to (0, -36.52, 2.61) mm, rotated rx 27.76 ry 0 rz 180 deg; joints [15.756, -63.263, 106.951, -157.781, 45.898, 101.888]
  MoveL 4186 to (-200, -36.52, 2.61) mm, rotated rx 27.76 ry 0 rz 180 deg; joints [18.278, -74.049, 122.693, -156.249, 51.142, 102.324]
  MoveL 4187 to (-200, -35.98, 2.34) mm, rotated rx 25.3 ry 0 rz 180 deg; joints [18.664, -73.273, 122.82, -156.064, 52.07, 100.039]
  MoveL 4188 to (0, -35.98, 2.34) mm, rotated rx 25.3 ry 0 rz 180 deg; joints [16.095, -62.617, 107.058, -157.604, 46.687, 99.516]
  MoveL 4189 to (0, -35.44, 2.1) mm, rotated rx 22.85 ry 0 rz 180 deg; joints [16.41, -61.955, 107.168, -157.464, 47.486, 97.182]
  MoveL 4190 to (-200, -35.44, 2.1) mm, rotated rx 22.85 ry 0 rz 180 deg; joints [19.022, -72.477, 122.949, -155.916, 53.009, 97.793]
  MoveL 4191 to (-200, -34.88, 1.88) mm, rotated rx 20.39 ry 0 rz 180 deg; joints [19.353, -71.661, 123.081, -155.805, 53.958, 95.582]
  MoveL 4192 to (0, -34.88, 1.88) mm, rotated rx 20.39 ry 0 rz 180 deg; joints [16.701, -61.277, 107.281, -157.36, 48.294, 94.881]
  MoveL 4193 to (0, -34.31, 1.68) mm, rotated rx 17.93 ry 0 rz 180 deg; joints [16.968, -60.584, 107.395, -157.291, 49.11, 92.615]
  MoveL 4194 to (-200, -34.31, 1.68) mm, rotated rx 17.93 ry 0 rz 180 deg; joints [19.656, -70.828, 123.214, -155.728, 54.917, 93.405]
  MoveL 4195 to (-200, -33.74, 1.51) mm, rotated rx 15.48 ry 0 rz 180 deg; joints [19.931, -69.978, 123.349, -155.684, 55.882, 91.258]
  MoveL 4196 to (0, -33.74, 1.51) mm, rotated rx 15.48 ry 0 rz 180 deg; joints [17.211, -59.878, 107.512, -157.255, 49.932, 90.377]
  MoveL 4197 to (0, -33.16, 1.36) mm, rotated rx 13.02 ry 0 rz 180 deg; joints [17.428, -59.16, 107.629, -157.25, 50.759, 88.167]
  MoveL 4198 to (-200, -33.16, 1.36) mm, rotated rx 13.02 ry 0 rz 180 deg; joints [20.178, -69.112, 123.484, -155.671, 56.854, 89.138]
  MoveL 4199 to (-200, -32.57, 1.24) mm, rotated rx 10.57 ry 0 rz 180 deg; joints [20.396, -68.231, 123.619, -155.688, 57.831, 87.043]
  MoveL 4200 to (0, -32.57, 1.24) mm, rotated rx 10.57 ry 0 rz 180 deg; joints [17.621, -58.43, 107.748, -157.275, 51.591, 85.983]
  MoveL 4201 to (0, -31.98, 1.14) mm, rotated rx 8.11 ry 0 rz 180 deg; joints [17.788, -57.689, 107.866, -157.328, 52.425, 83.822]
  MoveL 4202 to (-200, -31.98, 1.14) mm, rotated rx 8.11 ry 0 rz 180 deg; joints [20.585, -67.338, 123.753, -155.732, 58.812, 84.972]
  MoveL 4203 to (-200, -31.38, 1.07) mm, rotated rx 5.66 ry 0 rz 180 deg; joints [20.746, -66.433, 123.887, -155.804, 59.796, 82.919]
  MoveL 4204 to (0, -31.38, 1.07) mm, rotated rx 5.66 ry 0 rz 180 deg; joints [17.93, -56.94, 107.985, -157.409, 53.261, 81.681]
  MoveL 4205 to (0, -30.78, 1.02) mm, rotated rx 3.2 ry 0 rz 180 deg; joints [18.046, -56.182, 108.104, -157.516, 54.098, 79.56]
  MoveL 4206 to (-200, -30.78, 1.02) mm, rotated rx 3.2 ry 0 rz 180 deg; joints [20.877, -65.517, 124.02, -155.901, 60.781, 80.885]
  MoveL 4207 to (-200, -30.18, 1) mm, rotated rx 0.75 ry 0 rz 180 deg; joints [20.979, -64.592, 124.151, -156.022, 61.767, 78.864]
  MoveL 4208 to (0, -30.18, 1) mm, rotated rx 0.75 ry 0 rz 180 deg; joints [18.136, -55.417, 108.221, -157.647, 54.935, 77.454]
  MoveL 4209 to (0, -29.58, 1) mm, rotated rx 0 ry 0 rz 180 deg; joints [18.159, -55.165, 108.261, -157.698, 55.211, 76.829]
  MoveL 4210 to (-200, -29.58, 1) mm, rotated rx 0 ry 0 rz 180 deg; joints [21.005, -64.286, 124.195, -156.07, 62.092, 78.266]
  MoveL 4211 to (-200, -28.98, 1) mm, rotated rx 0 ry 0 rz 180 deg; joints [21.005, -64.252, 124.202, -156.079, 62.129, 78.285]
  MoveL 4212 to (0, -28.98, 1) mm, rotated rx 0 ry 0 rz 180 deg; joints [18.159, -55.137, 108.268, -157.707, 55.242, 76.844]
  MoveL 4213 to (0, -28.38, 1) mm, rotated rx 0 ry 0 rz 180 deg; joints [18.159, -55.109, 108.274, -157.716, 55.274, 76.86]
  MoveL 4214 to (-200, -28.38, 1) mm, rotated rx 0 ry 0 rz 180 deg; joints [21.005, -64.218, 124.209, -156.088, 62.167, 78.304]
  MoveL 4215 to (-200, -27.78, 1) mm, rotated rx 0 ry 0 rz 180 deg; joints [21.005, -64.184, 124.216, -156.096, 62.204, 78.322]
  MoveL 4216 to (0, -27.78, 1) mm, rotated rx 0 ry 0 rz 180 deg; joints [18.159, -55.081, 108.28, -157.725, 55.306, 76.876]
  MoveL 4217 to (0, -27.18, 1) mm, rotated rx 0 ry 0 rz 180 deg; joints [18.159, -55.053, 108.286, -157.734, 55.337, 76.892]
  MoveL 4218 to (-200, -27.18, 1) mm, rotated rx 0 ry 0 rz 180 deg; joints [21.005, -64.15, 124.223, -156.105, 62.241, 78.341]
  MoveL 4219 to (-200, -26.58, 1) mm, rotated rx 0 ry 0 rz 180 deg; joints [21.005, -64.116, 124.229, -156.114, 62.278, 78.36]
  MoveL 4220 to (0, -26.58, 1) mm, rotated rx 0 ry 0 rz 180 deg; joints [18.159, -55.025, 108.293, -157.743, 55.369, 76.907]
  MoveL 4221 to (0, -25.98, 1) mm, rotated rx 0 ry 0 rz 180 deg; joints [18.159, -54.997, 108.299, -157.752, 55.401, 76.923]
  MoveL 4222 to (-200, -25.98, 1) mm, rotated rx 0 ry 0 rz 180 deg; joints [21.005, -64.082, 124.236, -156.122, 62.316, 78.378]
  MoveL 4223 to (-200, -25.38, 1) mm, rotated rx 0 ry 0 rz 180 deg; joints [21.005, -64.048, 124.243, -156.131, 62.353, 78.397]
  MoveL 4224 to (0, -25.38, 1) mm, rotated rx 0 ry 0 rz 180 deg; joints [18.159, -54.969, 108.305, -157.761, 55.432, 76.939]
  MoveL 4225 to (0, -24.78, 1) mm, rotated rx 0 ry 0 rz 180 deg; joints [18.159, -54.941, 108.311, -157.77, 55.464, 76.955]
  MoveL 4226 to (-200, -24.78, 1) mm, rotated rx 0 ry 0 rz 180 deg; joints [21.005, -64.014, 124.249, -156.14, 62.39, 78.415]
  MoveL 4227 to (-200, -24.18, 1) mm, rotated rx 0 ry 0 rz 180 deg; joints [21.005, -63.98, 124.256, -156.148, 62.427, 78.434]
  MoveL 4228 to (0, -24.18, 1) mm, rotated rx 0 ry 0 rz 180 deg; joints [18.159, -54.913, 108.317, -157.779, 55.495, 76.97]
  MoveL 4229 to (0, -23.58, 1) mm, rotated rx 0 ry 0 rz 180 deg; joints [18.159, -54.885, 108.323, -157.788, 55.527, 76.986]
  MoveL 4230 to (-200, -23.58, 1) mm, rotated rx 0 ry 0 rz 180 deg; joints [21.005, -63.946, 124.263, -156.157, 62.464, 78.453]
  MoveL 4231 to (-200, -22.98, 1) mm, rotated rx 0 ry 0 rz 180 deg; joints [21.005, -63.912, 124.269, -156.165, 62.502, 78.471]
  MoveL 4232 to (0, -22.98, 1) mm, rotated rx 0 ry 0 rz 180 deg; joints [18.159, -54.857, 108.329, -157.797, 55.559, 77.002]
  MoveL 4233 to (0, -22.38, 1) mm, rotated rx 0 ry 0 rz 180 deg; joints [18.159, -54.828, 108.335, -157.806, 55.59, 77.017]
  MoveL 4234 to (-200, -22.38, 1) mm, rotated rx 0 ry 0 rz 180 deg; joints [21.005, -63.878, 124.276, -156.174, 62.539, 78.49]
  MoveL 4235 to (-200, -21.78, 1) mm, rotated rx 0 ry 0 rz 180 deg; joints [21.005, -63.843, 124.282, -156.182, 62.576, 78.508]
  MoveL 4236 to (0, -21.78, 1) mm, rotated rx 0 ry 0 rz 180 deg; joints [18.159, -54.8, 108.341, -157.814, 55.622, 77.033]
  MoveL 4237 to (0, -21.18, 1) mm, rotated rx 0 ry 0 rz 180 deg; joints [18.159, -54.772, 108.347, -157.823, 55.653, 77.048]
  MoveL 4238 to (-200, -21.18, 1) mm, rotated rx 0 ry 0 rz 180 deg; joints [21.005, -63.809, 124.289, -156.191, 62.613, 78.527]
  MoveL 4239 to (-200, -20.58, 1) mm, rotated rx 0 ry 0 rz 180 deg; joints [21.005, -63.775, 124.295, -156.199, 62.65, 78.545]
  MoveL 4240 to (0, -20.58, 1) mm, rotated rx 0 ry 0 rz 180 deg; joints [18.159, -54.744, 108.353, -157.832, 55.685, 77.064]
  MoveL 4241 to (0, -19.98, 1) mm, rotated rx 0 ry 0 rz 180 deg; joints [18.159, -54.716, 108.359, -157.841, 55.716, 77.08]
  MoveL 4242 to (-200, -19.98, 1) mm, rotated rx 0 ry 0 rz 180 deg; joints [21.005, -63.741, 124.301, -156.208, 62.687, 78.564]
  MoveL 4243 to (-200, -19.38, 1) mm, rotated rx 0 ry 0 rz 180 deg; joints [21.005, -63.706, 124.308, -156.216, 62.725, 78.582]
  MoveL 4244 to (0, -19.38, 1) mm, rotated rx 0 ry 0 rz 180 deg; joints [18.159, -54.688, 108.365, -157.849, 55.748, 77.095]
  MoveL 4245 to (0, -18.78, 1) mm, rotated rx 0 ry 0 rz 180 deg; joints [18.159, -54.659, 108.371, -157.858, 55.779, 77.111]
  MoveL 4246 to (-200, -18.78, 1) mm, rotated rx 0 ry 0 rz 180 deg; joints [21.005, -63.672, 124.314, -156.225, 62.762, 78.6]
  MoveL 4247 to (-200, -18.18, 1) mm, rotated rx 0 ry 0 rz 180 deg; joints [21.005, -63.638, 124.32, -156.233, 62.799, 78.619]
  MoveL 4248 to (0, -18.18, 1) mm, rotated rx 0 ry 0 rz 180 deg; joints [18.159, -54.631, 108.376, -157.867, 55.811, 77.126]
  MoveL 4249 to (0, -17.58, 1) mm, rotated rx 0 ry 0 rz 180 deg; joints [18.159, -54.603, 108.382, -157.876, 55.843, 77.142]
  MoveL 4250 to (-200, -17.58, 1) mm, rotated rx 0 ry 0 rz 180 deg; joints [21.005, -63.604, 124.326, -156.242, 62.836, 78.637]
  MoveL 4251 to (-200, -16.98, 1) mm, rotated rx 0 ry 0 rz 180 deg; joints [21.005, -63.569, 124.333, -156.25, 62.873, 78.656]
  MoveL 4252 to (0, -16.98, 1) mm, rotated rx 0 ry 0 rz 180 deg; joints [18.159, -54.575, 108.388, -157.884, 55.874, 77.157]
  MoveL 4253 to (0, -16.38, 1) mm, rotated rx 0 ry 0 rz 180 deg; joints [18.159, -54.546, 108.393, -157.893, 55.906, 77.172]
  MoveL 4254 to (-200, -16.38, 1) mm, rotated rx 0 ry 0 rz 180 deg; joints [21.005, -63.535, 124.339, -156.258, 62.91, 78.674]
  MoveL 4255 to (-200, -15.78, 1) mm, rotated rx 0 ry 0 rz 180 deg; joints [21.005, -63.5, 124.345, -156.267, 62.947, 78.692]
  MoveL 4256 to (0, -15.78, 1) mm, rotated rx 0 ry 0 rz 180 deg; joints [18.159, -54.518, 108.399, -157.902, 55.937, 77.188]
  MoveL 4257 to (0, -15.18, 1) mm, rotated rx 0 ry 0 rz 180 deg; joints [18.159, -54.49, 108.405, -157.91, 55.968, 77.203]
  MoveL 4258 to (-200, -15.18, 1) mm, rotated rx 0 ry 0 rz 180 deg; joints [21.005, -63.466, 124.351, -156.275, 62.985, 78.71]
  MoveL 4259 to (-200, -14.58, 1) mm, rotated rx 0 ry 0 rz 180 deg; joints [21.005, -63.432, 124.357, -156.283, 63.022, 78.729]
  MoveL 4260 to (0, -14.58, 1) mm, rotated rx 0 ry 0 rz 180 deg; joints [18.159, -54.461, 108.41, -157.919, 56, 77.219]
  MoveL 4261 to (0, -13.98, 1) mm, rotated rx 0 ry 0 rz 180 deg; joints [18.159, -54.433, 108.416, -157.927, 56.031, 77.234]
  MoveL 4262 to (-200, -13.98, 1) mm, rotated rx 0 ry 0 rz 180 deg; joints [21.005, -63.397, 124.363, -156.292, 63.059, 78.747]
  MoveL 4263 to (-200, -13.38, 1) mm, rotated rx 0 ry 0 rz 180 deg; joints [21.005, -63.363, 124.369, -156.3, 63.096, 78.765]
  MoveL 4264 to (0, -13.38, 1) mm, rotated rx 0 ry 0 rz 180 deg; joints [18.159, -54.404, 108.422, -157.936, 56.063, 77.25]
  MoveL 4265 to (0, -12.78, 1) mm, rotated rx 0 ry 0 rz 180 deg; joints [18.159, -54.376, 108.427, -157.945, 56.094, 77.265]
  MoveL 4266 to (-200, -12.78, 1) mm, rotated rx 0 ry 0 rz 180 deg; joints [21.005, -63.328, 124.375, -156.308, 63.133, 78.784]
  MoveL 4267 to (-200, -12.18, 1) mm, rotated rx 0 ry 0 rz 180 deg; joints [21.005, -63.294, 124.381, -156.316, 63.17, 78.802]
  MoveL 4268 to (0, -12.18, 1) mm, rotated rx 0 ry 0 rz 180 deg; joints [18.159, -54.348, 108.433, -157.953, 56.126, 77.28]
  MoveL 4269 to (0, -11.58, 1) mm, rotated rx 0 ry 0 rz 180 deg; joints [18.159, -54.319, 108.438, -157.962, 56.157, 77.296]
  MoveL 4270 to (-200, -11.58, 1) mm, rotated rx 0 ry 0 rz 180 deg; joints [21.005, -63.259, 124.387, -156.325, 63.207, 78.82]
  MoveL 4271 to (-200, -10.98, 1) mm, rotated rx 0 ry 0 rz 180 deg; joints [21.005, -63.225, 124.393, -156.333, 63.244, 78.838]
  MoveL 4272 to (0, -10.98, 1) mm, rotated rx 0 ry 0 rz 180 deg; joints [18.159, -54.291, 108.443, -157.97, 56.189, 77.311]
  MoveL 4273 to (0, -10.38, 1) mm, rotated rx 0 ry 0 rz 180 deg; joints [18.159, -54.262, 108.449, -157.979, 56.22, 77.326]
  MoveL 4274 to (-200, -10.38, 1) mm, rotated rx 0 ry 0 rz 180 deg; joints [21.005, -63.19, 124.399, -156.341, 63.281, 78.856]
  MoveL 4275 to (-200, -9.78, 1) mm, rotated rx 0 ry 0 rz 180 deg; joints [21.005, -63.155, 124.405, -156.349, 63.318, 78.875]
  MoveL 4276 to (0, -9.78, 1) mm, rotated rx 0 ry 0 rz 180 deg; joints [18.159, -54.234, 108.454, -157.987, 56.251, 77.341]
  MoveL 4277 to (0, -9.18, 1) mm, rotated rx 0 ry 0 rz 180 deg; joints [18.159, -54.205, 108.46, -157.996, 56.283, 77.357]
  MoveL 4278 to (-200, -9.18, 1) mm, rotated rx 0 ry 0 rz 180 deg; joints [21.005, -63.121, 124.411, -156.357, 63.355, 78.893]
  MoveL 4279 to (-200, -8.58, 1) mm, rotated rx 0 ry 0 rz 180 deg; joints [21.005, -63.086, 124.416, -156.365, 63.392, 78.911]
  MoveL 4280 to (0, -8.58, 1) mm, rotated rx 0 ry 0 rz 180 deg; joints [18.159, -54.177, 108.465, -158.004, 56.314, 77.372]
  MoveL 4281 to (0, -7.98, 1) mm, rotated rx 0 ry 0 rz 180 deg; joints [18.159, -54.148, 108.47, -158.013, 56.346, 77.387]
  MoveL 4282 to (-200, -7.98, 1) mm, rotated rx 0 ry 0 rz 180 deg; joints [21.005, -63.051, 124.422, -156.374, 63.429, 78.929]
  MoveL 4283 to (-200, -7.38, 1) mm, rotated rx 0 ry 0 rz 180 deg; joints [21.005, -63.017, 124.428, -156.382, 63.466, 78.947]
  MoveL 4284 to (0, -7.38, 1) mm, rotated rx 0 ry 0 rz 180 deg; joints [18.159, -54.12, 108.475, -158.021, 56.377, 77.402]
  MoveL 4285 to (0, -6.78, 1) mm, rotated rx 0 ry 0 rz 180 deg; joints [18.159, -54.091, 108.481, -158.029, 56.408, 77.418]
  MoveL 4286 to (-200, -6.78, 1) mm, rotated rx 0 ry 0 rz 180 deg; joints [21.005, -62.982, 124.434, -156.39, 63.503, 78.965]
  MoveL 4287 to (-200, -6.18, 1) mm, rotated rx 0 ry 0 rz 180 deg; joints [21.005, -62.947, 124.439, -156.398, 63.54, 78.983]
  MoveL 4288 to (0, -6.18, 1) mm, rotated rx 0 ry 0 rz 180 deg; joints [18.159, -54.062, 108.486, -158.038, 56.44, 77.433]
  MoveL 4289 to (0, -5.58, 1) mm, rotated rx 0 ry 0 rz 180 deg; joints [18.159, -54.034, 108.491, -158.046, 56.471, 77.448]
  MoveL 4290 to (-200, -5.58, 1) mm, rotated rx 0 ry 0 rz 180 deg; joints [21.005, -62.913, 124.445, -156.406, 63.577, 79.001]
  MoveL 4291 to (-200, -4.98, 1) mm, rotated rx 0 ry 0 rz 180 deg; joints [21.005, -62.878, 124.45, -156.414, 63.614, 79.019]
  MoveL 4292 to (0, -4.98, 1) mm, rotated rx 0 ry 0 rz 180 deg; joints [18.159, -54.005, 108.496, -158.055, 56.502, 77.463]
  MoveL 4293 to (0, -4.38, 1) mm, rotated rx 0 ry 0 rz 180 deg; joints [18.159, -53.977, 108.501, -158.063, 56.534, 77.478]
  MoveL 4294 to (-200, -4.38, 1) mm, rotated rx 0 ry 0 rz 180 deg; joints [21.005, -62.843, 124.456, -156.422, 63.651, 79.037]
  MoveL 4295 to (-200, -3.78, 1) mm, rotated rx 0 ry 0 rz 180 deg; joints [21.005, -62.808, 124.462, -156.43, 63.688, 79.055]
  MoveL 4296 to (0, -3.78, 1) mm, rotated rx 0 ry 0 rz 180 deg; joints [18.159, -53.948, 108.506, -158.071, 56.565, 77.493]
  MoveL 4297 to (0, -3.18, 1) mm, rotated rx 0 ry 0 rz 180 deg; joints [18.159, -53.919, 108.511, -158.08, 56.596, 77.508]
  MoveL 4298 to (-200, -3.18, 1) mm, rotated rx 0 ry 0 rz 180 deg; joints [21.005, -62.773, 124.467, -156.438, 63.725, 79.073]
  MoveL 4299 to (-200, -2.58, 1) mm, rotated rx 0 ry 0 rz 180 deg; joints [21.005, -62.738, 124.472, -156.446, 63.762, 79.091]
  MoveL 4300 to (0, -2.58, 1) mm, rotated rx 0 ry 0 rz 180 deg; joints [18.159, -53.891, 108.517, -158.088, 56.627, 77.523]
  MoveL 4301 to (0, -1.98, 1) mm, rotated rx 0 ry 0 rz 180 deg; joints [18.159, -53.862, 108.522, -158.096, 56.659, 77.538]
  MoveL 4302 to (-200, -1.98, 1) mm, rotated rx 0 ry 0 rz 180 deg; joints [21.005, -62.704, 124.478, -156.454, 63.799, 79.109]
  MoveL 4303 to (-200, -1.38, 1) mm, rotated rx 0 ry 0 rz 180 deg; joints [21.005, -62.669, 124.483, -156.462, 63.836, 79.127]
  MoveL 4304 to (0, -1.38, 1) mm, rotated rx 0 ry 0 rz 180 deg; joints [18.159, -53.833, 108.526, -158.104, 56.69, 77.554]
  MoveL 4305 to (0, -0.78, 1) mm, rotated rx 0 ry 0 rz 180 deg; joints [18.159, -53.804, 108.531, -158.113, 56.721, 77.569]
  MoveL 4306 to (-200, -0.78, 1) mm, rotated rx 0 ry 0 rz 180 deg; joints [21.005, -62.634, 124.489, -156.469, 63.873, 79.145]
  MoveL 4307 to (-200, -0.18, 1) mm, rotated rx 0 ry 0 rz 180 deg; joints [21.005, -62.599, 124.494, -156.477, 63.91, 79.163]
  MoveL 4308 to (0, -0.18, 1) mm, rotated rx 0 ry 0 rz 180 deg; joints [18.159, -53.776, 108.536, -158.121, 56.753, 77.584]
  MoveL 4309 to (0, 0, 1) mm, rotated rx 0 ry 0 rz 180 deg; joints [18.159, -53.767, 108.538, -158.123, 56.762, 77.588]
  MoveL 4310 to (-200, 0, 1) mm, rotated rx 0 ry 0 rz 180 deg; joints [21.005, -62.588, 124.496, -156.48, 63.921, 79.168]
  MoveL 4311 to (-200, 0, 0.6) mm, rotated rx 0 ry 0 rz 180 deg; joints [21.022, -62.582, 124.484, -156.46, 63.92, 79.158]
  MoveL 4312 to (0, 0, 0.6) mm, rotated rx 0 ry 0 rz 180 deg; joints [18.174, -53.761, 108.527, -158.105, 56.761, 77.576]
  MoveL 4313 to (0, -0.6, 0.6) mm, rotated rx 0 ry 0 rz 180 deg; joints [18.174, -53.79, 108.522, -158.096, 56.729, 77.561]
  MoveL 4314 to (-200, -0.6, 0.6) mm, rotated rx 0 ry 0 rz 180 deg; joints [21.022, -62.617, 124.479, -156.452, 63.883, 79.14]
  MoveL 4315 to (-200, -1.2, 0.6) mm, rotated rx 0 ry 0 rz 180 deg; joints [21.022, -62.652, 124.473, -156.444, 63.846, 79.122]
  MoveL 4316 to (0, -1.2, 0.6) mm, rotated rx 0 ry 0 rz 180 deg; joints [18.174, -53.818, 108.517, -158.088, 56.698, 77.546]
  MoveL 4317 to (0, -1.8, 0.6) mm, rotated rx 0 ry 0 rz 180 deg; joints [18.174, -53.847, 108.512, -158.08, 56.667, 77.531]
  MoveL 4318 to (-200, -1.8, 0.6) mm, rotated rx 0 ry 0 rz 180 deg; joints [21.022, -62.686, 124.468, -156.436, 63.809, 79.104]
  MoveL 4319 to (-200, -2.4, 0.6) mm, rotated rx 0 ry 0 rz 180 deg; joints [21.022, -62.721, 124.463, -156.428, 63.772, 79.086]
  MoveL 4320 to (0, -2.4, 0.6) mm, rotated rx 0 ry 0 rz 180 deg; joints [18.174, -53.876, 108.507, -158.071, 56.635, 77.516]
  MoveL 4321 to (0, -3, 0.6) mm, rotated rx 0 ry 0 rz 180 deg; joints [18.174, -53.904, 108.502, -158.063, 56.604, 77.501]
  MoveL 4322 to (-200, -3, 0.6) mm, rotated rx 0 ry 0 rz 180 deg; joints [21.022, -62.756, 124.457, -156.421, 63.735, 79.068]
  MoveL 4323 to (-200, -3.6, 0.6) mm, rotated rx 0 ry 0 rz 180 deg; joints [21.022, -62.791, 124.452, -156.413, 63.698, 79.05]
  MoveL 4324 to (0, -3.6, 0.6) mm, rotated rx 0 ry 0 rz 180 deg; joints [18.174, -53.933, 108.497, -158.055, 56.573, 77.486]
  MoveL 4325 to (0, -4.2, 0.6) mm, rotated rx 0 ry 0 rz 180 deg; joints [18.174, -53.962, 108.492, -158.047, 56.542, 77.471]
  MoveL 4326 to (-200, -4.2, 0.6) mm, rotated rx 0 ry 0 rz 180 deg; joints [21.022, -62.826, 124.446, -156.405, 63.661, 79.032]
  MoveL 4327 to (-200, -4.8, 0.6) mm, rotated rx 0 ry 0 rz 180 deg; joints [21.022, -62.861, 124.441, -156.397, 63.624, 79.014]
  MoveL 4328 to (0, -4.8, 0.6) mm, rotated rx 0 ry 0 rz 180 deg; joints [18.174, -53.99, 108.487, -158.038, 56.51, 77.456]
  MoveL 4329 to (0, -5.4, 0.6) mm, rotated rx 0 ry 0 rz 180 deg; joints [18.174, -54.019, 108.481, -158.03, 56.479, 77.44]
  MoveL 4330 to (-200, -5.4, 0.6) mm, rotated rx 0 ry 0 rz 180 deg; joints [21.022, -62.895, 124.435, -156.389, 63.587, 78.996]
  MoveL 4331 to (-200, -6, 0.6) mm, rotated rx 0 ry 0 rz 180 deg; joints [21.022, -62.93, 124.429, -156.381, 63.55, 78.978]
  MoveL 4332 to (0, -6, 0.6) mm, rotated rx 0 ry 0 rz 180 deg; joints [18.174, -54.048, 108.476, -158.021, 56.448, 77.425]
  MoveL 4333 to (0, -6.6, 0.6) mm, rotated rx 0 ry 0 rz 180 deg; joints [18.174, -54.076, 108.471, -158.013, 56.416, 77.41]
  MoveL 4334 to (-200, -6.6, 0.6) mm, rotated rx 0 ry 0 rz 180 deg; joints [21.022, -62.965, 124.424, -156.372, 63.513, 78.96]
  MoveL 4335 to (-200, -7.2, 0.6) mm, rotated rx 0 ry 0 rz 180 deg; joints [21.022, -63, 124.418, -156.364, 63.476, 78.942]
  MoveL 4336 to (0, -7.2, 0.6) mm, rotated rx 0 ry 0 rz 180 deg; joints [18.174, -54.105, 108.466, -158.005, 56.385, 77.395]
  MoveL 4337 to (0, -7.8, 0.6) mm, rotated rx 0 ry 0 rz 180 deg; joints [18.174, -54.133, 108.461, -157.996, 56.354, 77.38]
  MoveL 4338 to (-200, -7.8, 0.6) mm, rotated rx 0 ry 0 rz 180 deg; joints [21.022, -63.034, 124.412, -156.356, 63.439, 78.924]
  MoveL 4339 to (-200, -8.4, 0.6) mm, rotated rx 0 ry 0 rz 180 deg; joints [21.022, -63.069, 124.407, -156.348, 63.402, 78.906]
  MoveL 4340 to (0, -8.4, 0.6) mm, rotated rx 0 ry 0 rz 180 deg; joints [18.174, -54.162, 108.455, -157.988, 56.322, 77.364]
  MoveL 4341 to (0, -9, 0.6) mm, rotated rx 0 ry 0 rz 180 deg; joints [18.174, -54.191, 108.45, -157.979, 56.291, 77.349]
  MoveL 4342 to (-200, -9, 0.6) mm, rotated rx 0 ry 0 rz 180 deg; joints [21.022, -63.104, 124.401, -156.34, 63.365, 78.888]
  MoveL 4343 to (-200, -9.6, 0.6) mm, rotated rx 0 ry 0 rz 180 deg; joints [21.022, -63.138, 124.395, -156.332, 63.328, 78.869]
  MoveL 4344 to (0, -9.6, 0.6) mm, rotated rx 0 ry 0 rz 180 deg; joints [18.174, -54.219, 108.445, -157.971, 56.26, 77.334]
  MoveL 4345 to (0, -10.2, 0.6) mm, rotated rx 0 ry 0 rz 180 deg; joints [18.174, -54.248, 108.439, -157.962, 56.228, 77.319]
  MoveL 4346 to (-200, -10.2, 0.6) mm, rotated rx 0 ry 0 rz 180 deg; joints [21.022, -63.173, 124.389, -156.324, 63.291, 78.851]
  MoveL 4347 to (-200, -10.8, 0.6) mm, rotated rx 0 ry 0 rz 180 deg; joints [21.022, -63.207, 124.383, -156.316, 63.254, 78.833]
  MoveL 4348 to (0, -10.8, 0.6) mm, rotated rx 0 ry 0 rz 180 deg; joints [18.174, -54.276, 108.434, -157.954, 56.197, 77.303]
  MoveL 4349 to (0, -11.4, 0.6) mm, rotated rx 0 ry 0 rz 180 deg; joints [18.174, -54.305, 108.429, -157.945, 56.165, 77.288]
  MoveL 4350 to (-200, -11.4, 0.6) mm, rotated rx 0 ry 0 rz 180 deg; joints [21.022, -63.242, 124.378, -156.307, 63.217, 78.815]
  MoveL 4351 to (-200, -12, 0.6) mm, rotated rx 0 ry 0 rz 180 deg; joints [21.022, -63.277, 124.372, -156.299, 63.18, 78.797]
  MoveL 4352 to (0, -12, 0.6) mm, rotated rx 0 ry 0 rz 180 deg; joints [18.174, -54.333, 108.423, -157.937, 56.134, 77.273]
  MoveL 4353 to (0, -12.6, 0.6) mm, rotated rx 0 ry 0 rz 180 deg; joints [18.174, -54.361, 108.418, -157.928, 56.103, 77.257]
  MoveL 4354 to (-200, -12.6, 0.6) mm, rotated rx 0 ry 0 rz 180 deg; joints [21.022, -63.311, 124.366, -156.291, 63.143, 78.778]
  MoveL 4355 to (-200, -13.2, 0.6) mm, rotated rx 0 ry 0 rz 180 deg; joints [21.022, -63.346, 124.36, -156.283, 63.106, 78.76]
  MoveL 4356 to (0, -13.2, 0.6) mm, rotated rx 0 ry 0 rz 180 deg; joints [18.174, -54.39, 108.412, -157.92, 56.071, 77.242]
  MoveL 4357 to (0, -13.8, 0.6) mm, rotated rx 0 ry 0 rz 180 deg; joints [18.174, -54.418, 108.407, -157.911, 56.04, 77.227]
  MoveL 4358 to (-200, -13.8, 0.6) mm, rotated rx 0 ry 0 rz 180 deg; joints [21.022, -63.38, 124.354, -156.274, 63.069, 78.742]
  MoveL 4359 to (-200, -14.4, 0.6) mm, rotated rx 0 ry 0 rz 180 deg; joints [21.022, -63.414, 124.348, -156.266, 63.032, 78.724]
